{region 'Documentation'}
(*!
<summary>Number of occupied entries.</summary>
*)
{endregion}
{attribute 'monitoring' := 'call'}
PROPERTY PUBLIC ChildCount : UINT //! Number of occupied entries.
GET
ChildCount := FCount;
END_GET
END_PROPERTY

{region 'Documentation'}
(*!
<summary>Records the original array index and returns only registered entries; never invokes a child.</summary>
*)
{endregion}
METHOD PUBLIC GetChild : I_Orchestratable //! Copied child interface at the original occupied index; zero and a latched InvalidAccess for an invalid index.
VAR_INPUT
    Index : DINT; //! Original array index to record and resolve within the occupied prefix.
END_VAR
VAR
    Position : LINT;
END_VAR
GetChild := 0;
IF FReadCount < ReadCapacity THEN
    FReadCount := FReadCount + 1;
    FReadIndices[FReadCount] := Index;
ELSE
    FTraceOverflow := TRUE;
END_IF;

Position := DINT_TO_LINT(Index) - DINT_TO_LINT(FLowerBound) + 1;
IF (Position < 1) OR (Position > UINT_TO_LINT(FCount)) THEN
    FInvalidAccess := TRUE;
    RETURN;
END_IF;
GetChild := FChildren[LINT_TO_UINT(Position)];
END_METHOD

{region 'Documentation'}
(*!
<summary>Copies the fixed registered prefix and clears access evidence without retaining addresses.</summary>
*)
{endregion}
METHOD PUBLIC Initialize : BOOL //! TRUE after copying a valid nonzero occupied prefix; FALSE leaves ChildCount zero.
VAR_INPUT
    Count : UINT; //! Occupied prefix length in 1..ChildCapacity; it must fit the supplied array.
END_VAR
VAR_IN_OUT
    Children : ARRAY[*] OF I_Orchestratable; //! Borrowed array whose occupied interface prefix is copied; keep the referenced children alive.
END_VAR
VAR
    Position : UINT;
    ArrayIndex : DINT;
END_VAR
Initialize := FALSE;
FCount := 0;
FLowerBound := LOWER_BOUND(Children, 1);
FUpperBound := UPPER_BOUND(Children, 1);
FReadCount := 0;
FInvalidAccess := FALSE;
FTraceOverflow := FALSE;
FOR Position := 1 TO ChildCapacity DO
    FChildren[Position] := 0;
END_FOR;
FOR Position := 1 TO ReadCapacity DO
    FReadIndices[Position] := 0;
END_FOR;
IF (Count = 0) OR (Count > ChildCapacity)
    OR (DINT_TO_LINT(FLowerBound) + UINT_TO_LINT(Count) - 1 > DINT_TO_LINT(FUpperBound)) THEN
    RETURN;
END_IF;

FOR Position := 1 TO Count DO
    ArrayIndex := FLowerBound + UINT_TO_DINT(Position) - 1;
    IF Children[ArrayIndex] = 0 THEN
        RETURN;
    END_IF;
    FChildren[Position] := Children[ArrayIndex];
END_FOR;
FCount := Count;
Initialize := TRUE;
END_METHOD

{region 'Documentation'}
(*!
<summary>Latched access outside the registered range.</summary>
*)
{endregion}
{attribute 'monitoring' := 'call'}
PROPERTY PUBLIC InvalidAccess : BOOL //! Latched access outside the registered range.
GET
InvalidAccess := FInvalidAccess;
END_GET
END_PROPERTY

{region 'Documentation'}
(*!
<summary>Number of retained index-access observations.</summary>
*)
{endregion}
{attribute 'monitoring' := 'call'}
PROPERTY PUBLIC ReadCount : UINT //! Number of retained index-access observations.
GET
ReadCount := FReadCount;
END_GET
END_PROPERTY

{region 'Documentation'}
(*!
<summary>Whether the bounded index trace was exhausted.</summary>
*)
{endregion}
{attribute 'monitoring' := 'call'}
PROPERTY PUBLIC TraceOverflow : BOOL //! Whether the bounded index trace was exhausted.
GET
TraceOverflow := FTraceOverflow;
END_GET
END_PROPERTY

END_FUNCTION_BLOCK

// ---- SelfTests/Helper/Orchestration/OrchestrationChildDouble.TcPOU
{region 'Documentation'}
(*!
<summary>Controllable I_Orchestratable boundary for isolated scheduler tests.</summary>
<description>

Stimulus versus commands

The scenario supplies the next ObservationInput at the child FB call after the helper.
Request methods only record invocations; they do not select states or run a copied lifecycle.
This permits independent, explicitly authored normal and exceptional responses.
BeginCycle clears call counters before the helper without changing the prior observation.

Reservation boundary

BeginCycle supplies this cycle's reservation responses, defaulting to Accepted.
Only Accepted sets one local marker; waiting and failure leave it unchanged.
No global publisher or reservation is changed.
The tests verify orchestration call order, not the real owner's budget calculation.
</description>
*)
{endregion}
FUNCTION_BLOCK OrchestrationChildDouble IMPLEMENTS I_Orchestratable
VAR_INPUT
    ObservationInput : ST_OrchestrationObservation; //! Scripted view accepted only when this concrete child body is called.
END_VAR
VAR
    FName : STRING(GVL_Constants.NameLength);
    FExecutionSlot : UINT;
    FInitialized : BOOL;
    FObservation : ST_OrchestrationObservation;
    FCalls : ST_OrchestrationCalls;
    FReservedEntryCount : UINT;
    FExecutionReservationResult : E_EventReservationResult := E_EventReservationResult.Accepted;
    FResetReservationResult : E_EventReservationResult := E_EventReservationResult.Accepted;
END_VAR
VAR CONSTANT
    ReservationMarker : UINT := 1;
END_VAR

FCalls.BodyCount := FCalls.BodyCount + 1;
FObservation := ObservationInput;

{region 'Documentation'}
(*!
<summary>Clears call evidence and supplies reservation responses; retains the prior child view and marker.</summary>
*)
{endregion}
METHOD PUBLIC BeginCycle
VAR_INPUT
    ExecutionReservationResult : E_EventReservationResult := E_EventReservationResult.Accepted; //! Execution admission response for this cycle; Accepted sets the local marker.
    ResetReservationResult : E_EventReservationResult := E_EventReservationResult.Accepted; //! Reset admission response for this cycle; Accepted sets the local marker.
END_VAR
VAR
    EmptyCalls : ST_OrchestrationCalls;
END_VAR
FCalls := EmptyCalls;
FExecutionReservationResult := ExecutionReservationResult;
FResetReservationResult := ResetReservationResult;
END_METHOD

{region 'Documentation'}
(*!
<summary>Interface-call evidence for the current fixture cycle.</summary>
*)
{endregion}
{attribute 'monitoring' := 'variable'}
PROPERTY PUBLIC Calls : ST_OrchestrationCalls //! Interface-call evidence for the current fixture cycle.
GET
Calls := FCalls;
END_GET
END_PROPERTY

{region 'Documentation'}
(*!
<summary>Registration slot retained independently of cyclic observations.</summary>
*)
{endregion}
{attribute 'monitoring' := 'call'}
PROPERTY PUBLIC ExecutionSlot : UINT //! Registration slot retained independently of cyclic observations.
GET
ExecutionSlot := FExecutionSlot;
END_GET
SET
FExecutionSlot := ExecutionSlot;
END_SET
END_PROPERTY

{region 'Documentation'}
(*!
<summary>Releases only the local marker and records the released amount; repeated calls are idempotent.</summary>
*)
{endregion}
METHOD PUBLIC FreeReservedEvents : BOOL //! Always TRUE after clearing the local marker; the call and released amount remain recorded.
FCalls.FreeCount := FCalls.FreeCount + 1;
FCalls.ReleasedEntryCount := FCalls.ReleasedEntryCount + FReservedEntryCount;
FReservedEntryCount := 0;
FreeReservedEvents := TRUE;
END_METHOD

{region 'Documentation'}
(*!
<summary>Scripted child failure classification.</summary>
*)
{endregion}
{attribute 'monitoring' := 'call'}
PROPERTY PUBLIC HasError : BOOL //! Scripted child failure classification.
GET
HasError := FObservation.Result = E_Result.Error;
END_GET
END_PROPERTY

{region 'Documentation'}
(*!
<summary>Resets the local interface double; it has no timers, publisher or production lifecycle.</summary>
*)
{endregion}
METHOD PUBLIC Initialize
VAR_INPUT
    Name : STRING(GVL_Constants.NameLength); //! Diagnostic child name retained by the fixture.
    Slot : UINT; //! Registered execution slot retained independently of scripted observations.
END_VAR
VAR
    EmptyCalls : ST_OrchestrationCalls;
    InitialView : ST_OrchestrationObservation;
END_VAR
FName := Name;
FExecutionSlot := Slot;
FObservation := InitialView;
FCalls := EmptyCalls;
FReservedEntryCount := 0;
FExecutionReservationResult := E_EventReservationResult.Accepted;
FResetReservationResult := E_EventReservationResult.Accepted;
FInitialized := TRUE;
END_METHOD

{region 'Documentation'}
(*!
<summary>Scripted terminal completion signal.</summary>
*)
{endregion}
{attribute 'monitoring' := 'call'}
PROPERTY PUBLIC IsComplete : BOOL //! Scripted terminal completion signal.
GET
IsComplete := FObservation.Complete;
END_GET
END_PROPERTY

{region 'Documentation'}
(*!
<summary>Whether the double has been explicitly configured.</summary>
*)
{endregion}
{attribute 'monitoring' := 'call'}
PROPERTY PUBLIC IsInitialized : BOOL //! Whether the double has been explicitly configured.
GET
IsInitialized := FInitialized;
END_GET
END_PROPERTY

{region 'Documentation'}
(*!
<summary>Scripted readiness, independent of helper requests.</summary>
*)
{endregion}
{attribute 'monitoring' := 'call'}
PROPERTY PUBLIC IsReady : BOOL //! Scripted readiness, independent of helper requests.
GET
IsReady := FObservation.Ready;
END_GET
END_PROPERTY

{region 'Documentation'}
(*!
<summary>Diagnostic child identity.</summary>
*)
{endregion}
{attribute 'monitoring' := 'variable'}
PROPERTY PUBLIC Name : STRING(GVL_Constants.NameLength) //! Diagnostic child identity.
GET
Name := FName;
END_GET
END_PROPERTY

{region 'Documentation'}
(*!
<summary>Current scripted snapshot; requests cannot change it.</summary>
*)
{endregion}
{attribute 'monitoring' := 'variable'}
PROPERTY PUBLIC Observation : ST_OrchestrationObservation //! Current scripted snapshot; requests cannot change it.
GET
Observation := FObservation;
END_GET
END_PROPERTY

{region 'Documentation'}
(*!
<summary>Records the Abort request without changing the scripted state.</summary>
*)
{endregion}
METHOD PUBLIC RequestAbort
FCalls.AbortCount := FCalls.AbortCount + 1;
END_METHOD

{region 'Documentation'}
(*!
<summary>Records the Reset request without changing the scripted state.</summary>
*)
{endregion}
METHOD PUBLIC RequestReset
FCalls.ResetCount := FCalls.ResetCount + 1;

FCalls.ResetWithoutReservation := FCalls.ResetWithoutReservation OR (FReservedEntryCount = 0);
END_METHOD

{region 'Documentation'}
(*!
<summary>Records the Start request without changing the scripted state.</summary>
*)
{endregion}
METHOD PUBLIC RequestStart
FCalls.StartCount := FCalls.StartCount + 1;
FCalls.StartWithoutReservation := FCalls.StartWithoutReservation OR (FReservedEntryCount = 0);
END_METHOD

{region 'Documentation'}
(*!
<summary>Local admission marker, not a global Event Buffer contribution.</summary>
*)
{endregion}
{attribute 'monitoring' := 'call'}
PROPERTY PUBLIC ReservedEntryCount : UINT //! Local admission marker, not a global Event Buffer contribution.
GET
ReservedEntryCount := FReservedEntryCount;
END_GET
END_PROPERTY

{region 'Documentation'}
(*!
<summary>Returns the scripted execution admission response; only Accepted sets the local marker.</summary>
*)
{endregion}
METHOD PUBLIC ReserveExecutionEvents : E_EventReservationResult //! Scripted execution admission response; only Accepted installs the local marker.
FCalls.ExecutionReservationCount := FCalls.ExecutionReservationCount + 1;
IF FExecutionReservationResult = E_EventReservationResult.Accepted THEN
    FReservedEntryCount := ReservationMarker;
END_IF;
ReserveExecutionEvents := FExecutionReservationResult;
END_METHOD

{region 'Documentation'}
(*!
<summary>Returns the scripted reset admission response; only Accepted sets the local marker.</summary>
*)
{endregion}
METHOD PUBLIC ReserveResetEvents : E_EventReservationResult //! Scripted Reset admission response; only Accepted installs the local marker.
FCalls.ResetReservationCount := FCalls.ResetReservationCount + 1;
IF FResetReservationResult = E_EventReservationResult.Accepted THEN
    FReservedEntryCount := ReservationMarker;
END_IF;
ReserveResetEvents := FResetReservationResult;
END_METHOD

{region 'Documentation'}
(*!
<summary>Scripted child result.</summary>
*)
{endregion}
{attribute 'monitoring' := 'call'}
PROPERTY PUBLIC Result : E_Result //! Scripted child result.
GET
Result := FObservation.Result;
END_GET
END_PROPERTY

{region 'Documentation'}
(*!
<summary>View applied on the most recent child call.</summary>
*)
{endregion}
{attribute 'monitoring' := 'call'}
PROPERTY PUBLIC State : E_State //! View applied on the most recent child call.
GET
State := FObservation.State;
END_GET
END_PROPERTY

END_FUNCTION_BLOCK

// ---- SelfTests/TestCases/TestSuite_Orchestrator/Test_OrchestratorNegativeBounds.TcPOU
{region 'Documentation'}
(*!
<summary>Checks the same execution trace with actual indices -3 through -1.</summary>
*)
{endregion}
FUNCTION_BLOCK Test_OrchestratorNegativeBounds EXTENDS OrchestrationTestBase

SUPER^();

{region 'Documentation'}
(*!
<summary>Defines this scenario independently of the subject's internal fields.</summary>
*)
{endregion}
METHOD PROTECTED ConfigureScenario
FArrayLayout := E_OrchestrationArrayLayout.Negative;
FChildCount := 3;
ConfigureStandardSequence();
END_METHOD

END_FUNCTION_BLOCK

// ---- SelfTests/TestCases/TestSuite_Orchestrator/Test_OrchestratorUnusedCapacity.TcPOU
{region 'Documentation'}
(*!
<summary>Checks that unused array capacity at indices 4 through 6 is never processed.</summary>
*)
{endregion}
FUNCTION_BLOCK Test_OrchestratorUnusedCapacity EXTENDS OrchestrationTestBase

SUPER^();

{region 'Documentation'}
(*!
<summary>Defines this scenario independently of the subject's internal fields.</summary>
*)
{endregion}
METHOD PROTECTED ConfigureScenario
FArrayLayout := E_OrchestrationArrayLayout.SpareCapacity;
FChildCount := 3;
ConfigureStandardSequence();
END_METHOD

END_FUNCTION_BLOCK

// ---- SelfTests/TestCases/TestSuite_Orchestrator/Test_OrchestratorSingleChild.TcPOU
{region 'Documentation'}
(*!
<summary>Checks a single registered child without a successor or unused-capacity access.</summary>
*)
{endregion}
FUNCTION_BLOCK Test_OrchestratorSingleChild EXTENDS OrchestrationTestBase

SUPER^();

{region 'Documentation'}
(*!
<summary>Defines this scenario independently of the subject's internal fields.</summary>
*)
{endregion}
METHOD PROTECTED ConfigureScenario
FArrayLayout := E_OrchestrationArrayLayout.Ordinary;
FChildCount := 1;
FStepCount := 4;

{region "Cycle 01 - Idle readiness"}
FSteps[1].Task := E_OrchestratorTask.Idle;
FSteps[1].ExpectedReady := TRUE;
{endregion}

{region "Cycle 02 - Start child 1"}
FSteps[2].Children[1].State := E_State.Completed;
FSteps[2].Children[1].Ready := FALSE;
FSteps[2].Children[1].Complete := TRUE;
FSteps[2].Children[1].Result := E_Result.Passed;
FSteps[2].ExpectedStartChild := 1;
FSteps[2].ExpectedSlot := 1;
FSteps[2].ExpectedReservations[1] := 1;
{endregion}

{region "Cycle 03 - Completed observation"}
FSteps[3].Children[1].State := E_State.Completed;
FSteps[3].Children[1].Ready := FALSE;
FSteps[3].Children[1].Complete := TRUE;
FSteps[3].Children[1].Result := E_Result.Passed;
FSteps[3].ExpectedReleasedEntries[1] := 1;
FSteps[3].ExpectedFinished := TRUE;
{endregion}

{region "Cycle 04 - Completed observation"}
FSteps[4].Children[1].State := E_State.Completed;
FSteps[4].Children[1].Ready := FALSE;
FSteps[4].Children[1].Complete := TRUE;
FSteps[4].Children[1].Result := E_Result.Passed;
FSteps[4].ExpectedFinished := TRUE;
{endregion}
END_METHOD

END_FUNCTION_BLOCK

// ---- SelfTests/TestCases/TestSuite_Orchestrator/Test_OrchestratorIdleReadiness.TcPOU
{region 'Documentation'}
(*!
<summary>Checks that readiness follows prior child observations and recovers without dispatch or diagnostics.</summary>
*)
{endregion}
FUNCTION_BLOCK Test_OrchestratorIdleReadiness EXTENDS OrchestrationTestBase

SUPER^();

{region 'Documentation'}
(*!
<summary>Defines independent stimuli and expected requests, reservations, task status and diagnostic counts.</summary>
*)
{endregion}
METHOD PROTECTED ConfigureScenario
FStepCount := 4;

{region "01 - Make the second child not ready after helper observation"}
FSteps[1].Task := E_OrchestratorTask.Idle;
FSteps[1].Children[2].Ready := FALSE;
FSteps[1].ExpectedReady := TRUE;
{endregion}

{region "02 - Observe not-ready child without dispatch"}
FSteps[2].Task := E_OrchestratorTask.Idle;
FSteps[2].Children[2].Ready := FALSE;
{endregion}

{region "03 - Restore child readiness after this observation"}
FSteps[3].Task := E_OrchestratorTask.Idle;
{endregion}

{region "04 - Observe restored readiness"}
FSteps[4].Task := E_OrchestratorTask.Idle;
FSteps[4].ExpectedReady := TRUE;
{endregion}
END_METHOD

END_FUNCTION_BLOCK

// ---- SelfTests/TestCases/TestSuite_Orchestrator/Test_OrchestratorMissingStartReaction.TcPOU
{region 'Documentation'}
(*!
<summary>Detects missing Start response on the following call, releases its reservation and prevents retries.</summary>
*)
{endregion}
FUNCTION_BLOCK Test_OrchestratorMissingStartReaction EXTENDS OrchestrationTestBase

SUPER^();

{region 'Documentation'}
(*!
<summary>Defines independent stimuli and expected requests, reservations, task status and diagnostic counts.</summary>
*)
{endregion}
METHOD PROTECTED ConfigureScenario
FStepCount := 12;

{region "01 - Idle readiness before child processing"}
FSteps[1].Task := E_OrchestratorTask.Idle;
FSteps[1].ExpectedReady := TRUE;
{endregion}

{region "02 - Request Start but leave child Idle"}
FSteps[2].ExpectedStartChild := 1;
FSteps[2].ExpectedSlot := 1;
FSteps[2].ExpectedReservations[1] := 1;
{endregion}

{region "03 - Following helper call must reject missing response"}
FSteps[3].ExpectedSlot := 1;
FSteps[3].ExpectedDiagnosticCount := 1;
FSteps[3].ExpectedReleasedEntries[1] := 1;
FSteps[3].ExpectedResult := E_Result.Error;
{endregion}

{region "04 - No retry or duplicate diagnostic"}
FSteps[4].ExpectedSlot := 1;
FSteps[4].ExpectedDiagnosticCount := 1;
FSteps[4].ExpectedResult := E_Result.Error;
{endregion}

{region "05 - Idle preserves the held error"}
FSteps[5].Task := E_OrchestratorTask.Idle;
FSteps[5].ExpectedDiagnosticCount := 1;
FSteps[5].ExpectedResult := E_Result.Error;
{endregion}

{region "06 - Execution cannot bypass held error"}
FSteps[6].ExpectedDiagnosticCount := 1;
FSteps[6].ExpectedResult := E_Result.Error;
{endregion}

{region "07 - New Reset clears helper error without clearing captured evidence"}
FSteps[7].Task := E_OrchestratorTask.Reset;
FSteps[7].ExpectedDiagnosticCount := 1;
{endregion}

{region "08 - All already-ready children count as reset-complete"}
FSteps[8].Task := E_OrchestratorTask.Reset;
FSteps[8].ExpectedDiagnosticCount := 1;
FSteps[8].ExpectedResetFinished := TRUE;
{endregion}

{region "09 - Owner returns to ready Idle"}
FSteps[9].Task := E_OrchestratorTask.Idle;
FSteps[9].ExpectedDiagnosticCount := 1;
FSteps[9].ExpectedReady := TRUE;
{endregion}

{region "10 - Start is admitted again only after Reset"}
FSteps[10].Children[1].State := E_State.Completed;
FSteps[10].Children[1].Result := E_Result.Passed;
FSteps[10].Children[1].Ready := FALSE;
FSteps[10].Children[1].Complete := TRUE;
FSteps[10].ExpectedStartChild := 1;
FSteps[10].ExpectedSlot := 1;
FSteps[10].ExpectedDiagnosticCount := 1;
FSteps[10].ExpectedReservations[1] := 1;
{endregion}

{region "11 - Successful start response does not create another diagnostic"}
FSteps[11].Children[1].State := E_State.Completed;
FSteps[11].Children[1].Result := E_Result.Passed;
FSteps[11].Children[1].Ready := FALSE;
FSteps[11].Children[1].Complete := TRUE;
FSteps[11].ExpectedSlot := 2;
FSteps[11].ExpectedDiagnosticCount := 1;
FSteps[11].ExpectedReleasedEntries[1] := 1;
{endregion}

{region "12 - Owner stops the local scenario without starting later children"}
FSteps[12].Task := E_OrchestratorTask.Idle;
FSteps[12].Children[1].State := E_State.Completed;
FSteps[12].Children[1].Result := E_Result.Passed;
FSteps[12].Children[1].Ready := FALSE;
FSteps[12].Children[1].Complete := TRUE;
FSteps[12].ExpectedDiagnosticCount := 1;
{endregion}
END_METHOD

END_FUNCTION_BLOCK

// ---- SelfTests/TestCases/TestSuite_Orchestrator/Test_OrchestratorChildError.TcPOU
{region 'Documentation'}
(*!
<summary>Holds a child Error, prevents subsequent Starts and releases only after terminal observation.</summary>
*)
{endregion}
FUNCTION_BLOCK Test_OrchestratorChildError EXTENDS OrchestrationTestBase

SUPER^();

{region 'Documentation'}
(*!
<summary>Defines independent stimuli and expected requests, reservations, task status and diagnostic counts.</summary>
*)
{endregion}
METHOD PROTECTED ConfigureScenario
FStepCount := 8;

{region "01 - Idle readiness before child processing"}
FSteps[1].Task := E_OrchestratorTask.Idle;
FSteps[1].ExpectedReady := TRUE;
{endregion}

{region "02 - Start first child"}
FSteps[2].Children[1].State := E_State.Running;
FSteps[2].Children[1].Ready := FALSE;
FSteps[2].ExpectedStartChild := 1;
FSteps[2].ExpectedSlot := 1;
FSteps[2].ExpectedReservations[1] := 1;
{endregion}

{region "03 - Child reports Error after helper call"}
FSteps[3].Children[1].State := E_State.Running;
FSteps[3].Children[1].Result := E_Result.Error;
FSteps[3].Children[1].Ready := FALSE;
FSteps[3].ExpectedSlot := 1;
FSteps[3].ExpectedReservations[1] := 1;
{endregion}

{region "04 - Observe Error and retain active reservation"}
FSteps[4].Children[1].State := E_State.Running;
FSteps[4].Children[1].Result := E_Result.Error;
FSteps[4].Children[1].Ready := FALSE;
FSteps[4].ExpectedSlot := 1;
FSteps[4].ExpectedDiagnosticCount := 1;
FSteps[4].ExpectedReservations[1] := 1;
FSteps[4].ExpectedResult := E_Result.Error;
{endregion}

{region "05 - Failing child reaches terminal state"}
FSteps[5].Children[1].State := E_State.Completed;
FSteps[5].Children[1].Result := E_Result.Error;
FSteps[5].Children[1].Ready := FALSE;
FSteps[5].Children[1].Complete := TRUE;
FSteps[5].ExpectedSlot := 1;
FSteps[5].ExpectedDiagnosticCount := 1;
FSteps[5].ExpectedReservations[1] := 1;
FSteps[5].ExpectedResult := E_Result.Error;
{endregion}

{region "06 - Release terminal reservation without advancing execution"}
FSteps[6].Children[1].State := E_State.Completed;
FSteps[6].Children[1].Result := E_Result.Error;
FSteps[6].Children[1].Ready := FALSE;
FSteps[6].Children[1].Complete := TRUE;
FSteps[6].ExpectedSlot := 1;
FSteps[6].ExpectedDiagnosticCount := 1;
FSteps[6].ExpectedReleasedEntries[1] := 1;
FSteps[6].ExpectedResult := E_Result.Error;
{endregion}

{region "07 - Idle must not clear Error"}
FSteps[7].Task := E_OrchestratorTask.Idle;
FSteps[7].Children[1].State := E_State.Completed;
FSteps[7].Children[1].Result := E_Result.Error;
FSteps[7].Children[1].Ready := FALSE;
FSteps[7].Children[1].Complete := TRUE;
FSteps[7].ExpectedDiagnosticCount := 1;
FSteps[7].ExpectedResult := E_Result.Error;
{endregion}

{region "08 - Repeated Idle remains quiet"}
FSteps[8].Task := E_OrchestratorTask.Idle;
FSteps[8].Children[1].State := E_State.Completed;
FSteps[8].Children[1].Result := E_Result.Error;
FSteps[8].Children[1].Ready := FALSE;
FSteps[8].Children[1].Complete := TRUE;
FSteps[8].ExpectedDiagnosticCount := 1;
FSteps[8].ExpectedResult := E_Result.Error;
{endregion}
END_METHOD

END_FUNCTION_BLOCK

// ---- SelfTests/TestCases/TestSuite_Orchestrator/Test_OrchestratorUnexpectedAbort.TcPOU
{region 'Documentation'}
(*!
<summary>Treats a subordinate Abort during execution as a helper Error rather than normal completion.</summary>
*)
{endregion}
FUNCTION_BLOCK Test_OrchestratorUnexpectedAbort EXTENDS OrchestrationTestBase

SUPER^();

{region 'Documentation'}
(*!
<summary>Defines independent stimuli and expected requests, reservations, task status and diagnostic counts.</summary>
*)
{endregion}
METHOD PROTECTED ConfigureScenario
FStepCount := 6;

{region "01 - Idle readiness before child processing"}
FSteps[1].Task := E_OrchestratorTask.Idle;
FSteps[1].ExpectedReady := TRUE;
{endregion}

{region "02 - Start first child"}
FSteps[2].Children[1].State := E_State.Running;
FSteps[2].Children[1].Ready := FALSE;
FSteps[2].ExpectedStartChild := 1;
FSteps[2].ExpectedSlot := 1;
FSteps[2].ExpectedReservations[1] := 1;
{endregion}

{region "03 - Child reports unexpected Abort"}
FSteps[3].Children[1].State := E_State.Running;
FSteps[3].Children[1].Result := E_Result.Abort;
FSteps[3].Children[1].Ready := FALSE;
FSteps[3].ExpectedSlot := 1;
FSteps[3].ExpectedReservations[1] := 1;
{endregion}

{region "04 - Observe unexpected Abort while child finishes"}
FSteps[4].Children[1].State := E_State.Completed;
FSteps[4].Children[1].Result := E_Result.Abort;
FSteps[4].Children[1].Ready := FALSE;
FSteps[4].Children[1].Complete := TRUE;
FSteps[4].ExpectedSlot := 1;
FSteps[4].ExpectedDiagnosticCount := 1;
FSteps[4].ExpectedReservations[1] := 1;
FSteps[4].ExpectedResult := E_Result.Error;
{endregion}

{region "05 - Release without starting the successor"}
FSteps[5].Children[1].State := E_State.Completed;
FSteps[5].Children[1].Result := E_Result.Abort;
FSteps[5].Children[1].Ready := FALSE;
FSteps[5].Children[1].Complete := TRUE;
FSteps[5].ExpectedSlot := 1;
FSteps[5].ExpectedDiagnosticCount := 1;
FSteps[5].ExpectedReleasedEntries[1] := 1;
FSteps[5].ExpectedResult := E_Result.Error;
{endregion}

{region "06 - Held Error prevents a later Start"}
FSteps[6].Children[1].State := E_State.Completed;
FSteps[6].Children[1].Result := E_Result.Abort;
FSteps[6].Children[1].Ready := FALSE;
FSteps[6].Children[1].Complete := TRUE;
FSteps[6].ExpectedSlot := 1;
FSteps[6].ExpectedDiagnosticCount := 1;
FSteps[6].ExpectedResult := E_Result.Error;
{endregion}
END_METHOD

END_FUNCTION_BLOCK

// ---- SelfTests/TestCases/TestSuite_Orchestrator/Test_OrchestratorAbortInterruption.TcPOU
{region 'Documentation'}
(*!
<summary>Changes the owner task to Abort, requests only the active child and observes terminal cleanup.</summary>
*)
{endregion}
FUNCTION_BLOCK Test_OrchestratorAbortInterruption EXTENDS OrchestrationTestBase

SUPER^();

{region 'Documentation'}
(*!
<summary>Defines independent stimuli and expected requests, reservations, task status and diagnostic counts.</summary>
*)
{endregion}
METHOD PROTECTED ConfigureScenario
FStepCount := 8;

{region "01 - Idle readiness before child processing"}
FSteps[1].Task := E_OrchestratorTask.Idle;
FSteps[1].ExpectedReady := TRUE;
{endregion}

{region "02 - Start first child"}
FSteps[2].Children[1].State := E_State.Running;
FSteps[2].Children[1].Ready := FALSE;
FSteps[2].ExpectedStartChild := 1;
FSteps[2].ExpectedSlot := 1;
FSteps[2].ExpectedReservations[1] := 1;
{endregion}

{region "03 - Abort replaces Execution in the same helper call"}
FSteps[3].Task := E_OrchestratorTask.Abort;
FSteps[3].Children[1].State := E_State.Aborting;
FSteps[3].Children[1].Result := E_Result.Abort;
FSteps[3].Children[1].Ready := FALSE;
FSteps[3].ExpectedReservations[1] := 1;
FSteps[3].ExpectedAbortRequests[1] := 1;
{endregion}

{region "04 - Already-aborting child receives no duplicate request"}
FSteps[4].Task := E_OrchestratorTask.Abort;
FSteps[4].Children[1].State := E_State.Aborting;
FSteps[4].Children[1].Result := E_Result.Abort;
FSteps[4].Children[1].Ready := FALSE;
FSteps[4].ExpectedReservations[1] := 1;
{endregion}

{region "05 - Child reaches Completed with Abort"}
FSteps[5].Task := E_OrchestratorTask.Abort;
FSteps[5].Children[1].State := E_State.Completed;
FSteps[5].Children[1].Result := E_Result.Abort;
FSteps[5].Children[1].Ready := FALSE;
FSteps[5].Children[1].Complete := TRUE;
FSteps[5].ExpectedReservations[1] := 1;
{endregion}

{region "06 - Observe Abort completion and release"}
FSteps[6].Task := E_OrchestratorTask.Abort;
FSteps[6].Children[1].State := E_State.Completed;
FSteps[6].Children[1].Result := E_Result.Abort;
FSteps[6].Children[1].Ready := FALSE;
FSteps[6].Children[1].Complete := TRUE;
FSteps[6].ExpectedReleasedEntries[1] := 1;
FSteps[6].ExpectedAbortFinished := TRUE;
{endregion}

{region "07 - Completion does not select Idle autonomously"}
FSteps[7].Task := E_OrchestratorTask.Abort;
FSteps[7].Children[1].State := E_State.Completed;
FSteps[7].Children[1].Result := E_Result.Abort;
FSteps[7].Children[1].Ready := FALSE;
FSteps[7].Children[1].Complete := TRUE;
FSteps[7].ExpectedAbortFinished := TRUE;
{endregion}

{region "08 - Owner explicitly selects Idle"}
FSteps[8].Task := E_OrchestratorTask.Idle;
FSteps[8].Children[1].State := E_State.Completed;
FSteps[8].Children[1].Result := E_Result.Abort;
FSteps[8].Children[1].Ready := FALSE;
FSteps[8].Children[1].Complete := TRUE;
{endregion}
END_METHOD

END_FUNCTION_BLOCK

// ---- SelfTests/TestCases/TestSuite_Orchestrator/Test_OrchestratorIdleInterruption.TcPOU
{region 'Documentation'}
(*!
<summary>Idle stops new dispatch without forcing child Abort or releasing an unfinished reservation.</summary>
*)
{endregion}
FUNCTION_BLOCK Test_OrchestratorIdleInterruption EXTENDS OrchestrationTestBase

SUPER^();

{region 'Documentation'}
(*!
<summary>Defines independent stimuli and expected requests, reservations, task status and diagnostic counts.</summary>
*)
{endregion}
METHOD PROTECTED ConfigureScenario
FStepCount := 6;

{region "01 - Idle readiness before child processing"}
FSteps[1].Task := E_OrchestratorTask.Idle;
FSteps[1].ExpectedReady := TRUE;
{endregion}

{region "02 - Start first child"}
FSteps[2].Children[1].State := E_State.Running;
FSteps[2].Children[1].Ready := FALSE;
FSteps[2].ExpectedStartChild := 1;
FSteps[2].ExpectedSlot := 1;
FSteps[2].ExpectedReservations[1] := 1;
{endregion}

{region "03 - Idle leaves running child and reservation intact"}
FSteps[3].Task := E_OrchestratorTask.Idle;
FSteps[3].Children[1].State := E_State.Running;
FSteps[3].Children[1].Ready := FALSE;
FSteps[3].ExpectedReservations[1] := 1;
{endregion}

{region "04 - Child finishes while owner remains Idle"}
FSteps[4].Task := E_OrchestratorTask.Idle;
FSteps[4].Children[1].State := E_State.Completed;
FSteps[4].Children[1].Result := E_Result.Passed;
FSteps[4].Children[1].Ready := FALSE;
FSteps[4].Children[1].Complete := TRUE;
FSteps[4].ExpectedReservations[1] := 1;
{endregion}

{region "05 - Idle releases the finished child only"}
FSteps[5].Task := E_OrchestratorTask.Idle;
FSteps[5].Children[1].State := E_State.Completed;
FSteps[5].Children[1].Result := E_Result.Passed;
FSteps[5].Children[1].Ready := FALSE;
FSteps[5].Children[1].Complete := TRUE;
FSteps[5].ExpectedReleasedEntries[1] := 1;
{endregion}

{region "06 - Idle does not start the next child"}
FSteps[6].Task := E_OrchestratorTask.Idle;
FSteps[6].Children[1].State := E_State.Completed;
FSteps[6].Children[1].Result := E_Result.Passed;
FSteps[6].Children[1].Ready := FALSE;
FSteps[6].Children[1].Complete := TRUE;
{endregion}
END_METHOD

END_FUNCTION_BLOCK

// ---- SelfTests/TestCases/TestSuite_Orchestrator/Test_OrchestratorResetInterruption.TcPOU
{region 'Documentation'}
(*!
<summary>Reset replaces Execution and may dispatch subsequent child resets before prior reset completion.</summary>
*)
{endregion}
FUNCTION_BLOCK Test_OrchestratorResetInterruption EXTENDS OrchestrationTestBase

SUPER^();

{region 'Documentation'}
(*!
<summary>Defines independent stimuli and expected requests, reservations, task status and diagnostic counts.</summary>
*)
{endregion}
METHOD PROTECTED ConfigureScenario
FStepCount := 10;

{region "01 - Idle readiness before child processing"}
FSteps[1].Task := E_OrchestratorTask.Idle;
FSteps[1].ExpectedReady := TRUE;
{endregion}

{region "02 - Execution begins; other resources become not ready"}
FSteps[2].Children[1].State := E_State.Running;
FSteps[2].Children[1].Ready := FALSE;
FSteps[2].Children[2].Ready := FALSE;
FSteps[2].Children[3].Ready := FALSE;
FSteps[2].ExpectedStartChild := 1;
FSteps[2].ExpectedSlot := 1;
FSteps[2].ExpectedReservations[1] := 1;
{endregion}

{region "03 - Reset first child in the task-entry call"}
FSteps[3].Task := E_OrchestratorTask.Reset;
FSteps[3].Children[1].State := E_State.Reset;
FSteps[3].Children[1].Ready := FALSE;
FSteps[3].Children[2].Ready := FALSE;
FSteps[3].Children[3].Ready := FALSE;
FSteps[3].ExpectedResetChild := 1;
FSteps[3].ExpectedReservations[1] := 1;
{endregion}

{region "04 - Dispatch second Reset while first is still active"}
FSteps[4].Task := E_OrchestratorTask.Reset;
FSteps[4].Children[1].State := E_State.Reset;
FSteps[4].Children[1].Ready := FALSE;
FSteps[4].Children[2].State := E_State.Reset;
FSteps[4].Children[2].Ready := FALSE;
FSteps[4].Children[3].Ready := FALSE;
FSteps[4].ExpectedResetChild := 2;
FSteps[4].ExpectedReservations[1] := 1;
FSteps[4].ExpectedReservations[2] := 1;
{endregion}

{region "05 - Dispatch third Reset; first finishes afterwards"}
FSteps[5].Task := E_OrchestratorTask.Reset;
FSteps[5].Children[2].State := E_State.Reset;
FSteps[5].Children[2].Ready := FALSE;
FSteps[5].Children[3].State := E_State.Reset;
FSteps[5].Children[3].Ready := FALSE;
FSteps[5].ExpectedResetChild := 3;
FSteps[5].ExpectedReservations[1] := 1;
FSteps[5].ExpectedReservations[2] := 1;
FSteps[5].ExpectedReservations[3] := 1;
{endregion}

{region "06 - Release first; second finishes afterwards"}
FSteps[6].Task := E_OrchestratorTask.Reset;
FSteps[6].Children[3].State := E_State.Reset;
FSteps[6].Children[3].Ready := FALSE;
FSteps[6].ExpectedReservations[2] := 1;
FSteps[6].ExpectedReservations[3] := 1;
FSteps[6].ExpectedReleasedEntries[1] := 1;
{endregion}

{region "07 - Release second; third finishes afterwards"}
FSteps[7].Task := E_OrchestratorTask.Reset;
FSteps[7].ExpectedReservations[3] := 1;
FSteps[7].ExpectedReleasedEntries[2] := 1;
{endregion}

{region "08 - All reset observations are ready and reconciled"}
FSteps[8].Task := E_OrchestratorTask.Reset;
FSteps[8].ExpectedReleasedEntries[3] := 1;
FSteps[8].ExpectedResetFinished := TRUE;
{endregion}

{region "09 - Repeated Reset task does not restart dispatch"}
FSteps[9].Task := E_OrchestratorTask.Reset;
FSteps[9].ExpectedResetFinished := TRUE;
{endregion}

{region "10 - Only owner task change makes helper ready"}
FSteps[10].Task := E_OrchestratorTask.Idle;
FSteps[10].ExpectedReady := TRUE;
{endregion}
END_METHOD

END_FUNCTION_BLOCK

// ---- SelfTests/TestCases/TestSuite_Orchestrator/Test_OrchestratorResetContinuesAfterError.TcPOU
{region 'Documentation'}
(*!
<summary>Reset ignores unprocessed stale results, retains processed child errors and still attempts every child.</summary>
*)
{endregion}
FUNCTION_BLOCK Test_OrchestratorResetContinuesAfterError EXTENDS OrchestrationTestBase

SUPER^();

{region 'Documentation'}
(*!
<summary>Defines independent stimuli and expected requests, reservations, task status and diagnostic counts.</summary>
*)
{endregion}
METHOD PROTECTED ConfigureScenario
FStepCount := 8;

{region "01 - Establish previous terminal results through child calls"}
FSteps[1].Task := E_OrchestratorTask.Idle;
FSteps[1].Children[1].State := E_State.Completed;
FSteps[1].Children[1].Result := E_Result.Passed;
FSteps[1].Children[1].Ready := FALSE;
FSteps[1].Children[1].Complete := TRUE;
FSteps[1].Children[2].State := E_State.Completed;
FSteps[1].Children[2].Result := E_Result.Error;
FSteps[1].Children[2].Ready := FALSE;
FSteps[1].Children[2].Complete := TRUE;
FSteps[1].Children[3].State := E_State.Completed;
FSteps[1].Children[3].Result := E_Result.Passed;
FSteps[1].Children[3].Ready := FALSE;
FSteps[1].Children[3].Complete := TRUE;
FSteps[1].ExpectedReady := TRUE;
{endregion}

{region "02 - Reset first; ignore old Error in not-yet-reset second child"}
FSteps[2].Task := E_OrchestratorTask.Reset;
FSteps[2].Children[1].State := E_State.Completed;
FSteps[2].Children[1].Result := E_Result.Error;
FSteps[2].Children[1].Ready := FALSE;
FSteps[2].Children[1].Complete := TRUE;
FSteps[2].Children[2].State := E_State.Completed;
FSteps[2].Children[2].Result := E_Result.Error;
FSteps[2].Children[2].Ready := FALSE;
FSteps[2].Children[2].Complete := TRUE;
FSteps[2].Children[3].State := E_State.Completed;
FSteps[2].Children[3].Result := E_Result.Passed;
FSteps[2].Children[3].Ready := FALSE;
FSteps[2].Children[3].Complete := TRUE;
FSteps[2].ExpectedResetChild := 1;
FSteps[2].ExpectedReservations[1] := 1;
{endregion}

{region "03 - First Reset failed; still dispatch second"}
FSteps[3].Task := E_OrchestratorTask.Reset;
FSteps[3].Children[1].State := E_State.Completed;
FSteps[3].Children[1].Result := E_Result.Error;
FSteps[3].Children[1].Ready := FALSE;
FSteps[3].Children[1].Complete := TRUE;
FSteps[3].Children[2].State := E_State.Reset;
FSteps[3].Children[2].Ready := FALSE;
FSteps[3].Children[3].State := E_State.Completed;
FSteps[3].Children[3].Result := E_Result.Passed;
FSteps[3].Children[3].Ready := FALSE;
FSteps[3].Children[3].Complete := TRUE;
FSteps[3].ExpectedResetChild := 2;
FSteps[3].ExpectedDiagnosticCount := 1;
FSteps[3].ExpectedReservations[1] := 1;
FSteps[3].ExpectedReservations[2] := 1;
FSteps[3].ExpectedResult := E_Result.Error;
{endregion}

{region "04 - Keep failure while dispatching third"}
FSteps[4].Task := E_OrchestratorTask.Reset;
FSteps[4].Children[1].State := E_State.Completed;
FSteps[4].Children[1].Result := E_Result.Error;
FSteps[4].Children[1].Ready := FALSE;
FSteps[4].Children[1].Complete := TRUE;
FSteps[4].Children[3].State := E_State.Reset;
FSteps[4].Children[3].Ready := FALSE;
FSteps[4].ExpectedResetChild := 3;
FSteps[4].ExpectedDiagnosticCount := 1;
FSteps[4].ExpectedReservations[1] := 1;
FSteps[4].ExpectedReservations[2] := 1;
FSteps[4].ExpectedReservations[3] := 1;
FSteps[4].ExpectedResult := E_Result.Error;
{endregion}

{region "05 - Release successful second Reset"}
FSteps[5].Task := E_OrchestratorTask.Reset;
FSteps[5].Children[1].State := E_State.Completed;
FSteps[5].Children[1].Result := E_Result.Error;
FSteps[5].Children[1].Ready := FALSE;
FSteps[5].Children[1].Complete := TRUE;
FSteps[5].ExpectedDiagnosticCount := 1;
FSteps[5].ExpectedReservations[1] := 1;
FSteps[5].ExpectedReservations[3] := 1;
FSteps[5].ExpectedReleasedEntries[2] := 1;
FSteps[5].ExpectedResult := E_Result.Error;
{endregion}

{region "06 - Failed terminal child counts as finished, not ready"}
FSteps[6].Task := E_OrchestratorTask.Reset;
FSteps[6].Children[1].State := E_State.Completed;
FSteps[6].Children[1].Result := E_Result.Error;
FSteps[6].Children[1].Ready := FALSE;
FSteps[6].Children[1].Complete := TRUE;
FSteps[6].ExpectedDiagnosticCount := 1;
FSteps[6].ExpectedReservations[1] := 1;
FSteps[6].ExpectedReleasedEntries[3] := 1;
FSteps[6].ExpectedResetFinished := TRUE;
FSteps[6].ExpectedResult := E_Result.Error;
{endregion}

{region "07 - Idle reconciles failed terminal child reservation"}
FSteps[7].Task := E_OrchestratorTask.Idle;
FSteps[7].Children[1].State := E_State.Completed;
FSteps[7].Children[1].Result := E_Result.Error;
FSteps[7].Children[1].Ready := FALSE;
FSteps[7].Children[1].Complete := TRUE;
FSteps[7].ExpectedDiagnosticCount := 1;
FSteps[7].ExpectedReleasedEntries[1] := 1;
FSteps[7].ExpectedResult := E_Result.Error;
{endregion}

{region "08 - No additional diagnostic or dispatch in Idle"}
FSteps[8].Task := E_OrchestratorTask.Idle;
FSteps[8].Children[1].State := E_State.Completed;
FSteps[8].Children[1].Result := E_Result.Error;
FSteps[8].Children[1].Ready := FALSE;
FSteps[8].Children[1].Complete := TRUE;
FSteps[8].ExpectedDiagnosticCount := 1;
FSteps[8].ExpectedResult := E_Result.Error;
{endregion}
END_METHOD

END_FUNCTION_BLOCK

// ---- SelfTests/TestCases/TestSuite_Orchestrator/Test_OrchestratorRepeatAfterReset.TcPOU
{region 'Documentation'}
(*!
<summary>Runs all three children twice with intervening Reset and without reinitializing the subject or capture.</summary>
*)
{endregion}
FUNCTION_BLOCK Test_OrchestratorRepeatAfterReset EXTENDS OrchestrationTestBase

SUPER^();

{region 'Documentation'}
(*!
<summary>Defines independent stimuli and expected requests, reservations, task status and diagnostic counts.</summary>
*)
{endregion}
METHOD PROTECTED ConfigureScenario
FStepCount := 21;

{region "01 - Idle readiness before child processing"}
FSteps[1].Task := E_OrchestratorTask.Idle;
FSteps[1].ExpectedReady := TRUE;
{endregion}

{region "02 - First child completes on its Start call"}
FSteps[2].Children[1].State := E_State.Completed;
FSteps[2].Children[1].Result := E_Result.Passed;
FSteps[2].Children[1].Ready := FALSE;
FSteps[2].Children[1].Complete := TRUE;
FSteps[2].ExpectedStartChild := 1;
FSteps[2].ExpectedSlot := 1;
FSteps[2].ExpectedReservations[1] := 1;
{endregion}

{region "03 - Observe first completion"}
FSteps[3].Children[1].State := E_State.Completed;
FSteps[3].Children[1].Result := E_Result.Passed;
FSteps[3].Children[1].Ready := FALSE;
FSteps[3].Children[1].Complete := TRUE;
FSteps[3].ExpectedSlot := 2;
FSteps[3].ExpectedReleasedEntries[1] := 1;
{endregion}

{region "04 - Second child completes on its Start call"}
FSteps[4].Children[1].State := E_State.Completed;
FSteps[4].Children[1].Result := E_Result.Passed;
FSteps[4].Children[1].Ready := FALSE;
FSteps[4].Children[1].Complete := TRUE;
FSteps[4].Children[2].State := E_State.Completed;
FSteps[4].Children[2].Result := E_Result.Passed;
FSteps[4].Children[2].Ready := FALSE;
FSteps[4].Children[2].Complete := TRUE;
FSteps[4].ExpectedStartChild := 2;
FSteps[4].ExpectedSlot := 2;
FSteps[4].ExpectedReservations[2] := 1;
{endregion}

{region "05 - Observe second completion"}
FSteps[5].Children[1].State := E_State.Completed;
FSteps[5].Children[1].Result := E_Result.Passed;
FSteps[5].Children[1].Ready := FALSE;
FSteps[5].Children[1].Complete := TRUE;
FSteps[5].Children[2].State := E_State.Completed;
FSteps[5].Children[2].Result := E_Result.Passed;
FSteps[5].Children[2].Ready := FALSE;
FSteps[5].Children[2].Complete := TRUE;
FSteps[5].ExpectedSlot := 3;
FSteps[5].ExpectedReleasedEntries[2] := 1;
{endregion}

{region "06 - Third child completes on its Start call"}
FSteps[6].Children[1].State := E_State.Completed;
FSteps[6].Children[1].Result := E_Result.Passed;
FSteps[6].Children[1].Ready := FALSE;
FSteps[6].Children[1].Complete := TRUE;
FSteps[6].Children[2].State := E_State.Completed;
FSteps[6].Children[2].Result := E_Result.Passed;
FSteps[6].Children[2].Ready := FALSE;
FSteps[6].Children[2].Complete := TRUE;
FSteps[6].Children[3].State := E_State.Completed;
FSteps[6].Children[3].Result := E_Result.Passed;
FSteps[6].Children[3].Ready := FALSE;
FSteps[6].Children[3].Complete := TRUE;
FSteps[6].ExpectedStartChild := 3;
FSteps[6].ExpectedSlot := 3;
FSteps[6].ExpectedReservations[3] := 1;
{endregion}

{region "07 - Observe execution completion"}
FSteps[7].Children[1].State := E_State.Completed;
FSteps[7].Children[1].Result := E_Result.Passed;
FSteps[7].Children[1].Ready := FALSE;
FSteps[7].Children[1].Complete := TRUE;
FSteps[7].Children[2].State := E_State.Completed;
FSteps[7].Children[2].Result := E_Result.Passed;
FSteps[7].Children[2].Ready := FALSE;
FSteps[7].Children[2].Complete := TRUE;
FSteps[7].Children[3].State := E_State.Completed;
FSteps[7].Children[3].Result := E_Result.Passed;
FSteps[7].Children[3].Ready := FALSE;
FSteps[7].Children[3].Complete := TRUE;
FSteps[7].ExpectedReleasedEntries[3] := 1;
FSteps[7].ExpectedFinished := TRUE;
{endregion}

{region "08 - Completed Execution task is retained"}
FSteps[8].Children[1].State := E_State.Completed;
FSteps[8].Children[1].Result := E_Result.Passed;
FSteps[8].Children[1].Ready := FALSE;
FSteps[8].Children[1].Complete := TRUE;
FSteps[8].Children[2].State := E_State.Completed;
FSteps[8].Children[2].Result := E_Result.Passed;
FSteps[8].Children[2].Ready := FALSE;
FSteps[8].Children[2].Complete := TRUE;
FSteps[8].Children[3].State := E_State.Completed;
FSteps[8].Children[3].Result := E_Result.Passed;
FSteps[8].Children[3].Ready := FALSE;
FSteps[8].Children[3].Complete := TRUE;
FSteps[8].ExpectedFinished := TRUE;
{endregion}

{region "09 - Reset first completed child"}
FSteps[9].Task := E_OrchestratorTask.Reset;
FSteps[9].Children[2].State := E_State.Completed;
FSteps[9].Children[2].Result := E_Result.Passed;
FSteps[9].Children[2].Ready := FALSE;
FSteps[9].Children[2].Complete := TRUE;
FSteps[9].Children[3].State := E_State.Completed;
FSteps[9].Children[3].Result := E_Result.Passed;
FSteps[9].Children[3].Ready := FALSE;
FSteps[9].Children[3].Complete := TRUE;
FSteps[9].ExpectedResetChild := 1;
FSteps[9].ExpectedReservations[1] := 1;
{endregion}

{region "10 - Release first and Reset second"}
FSteps[10].Task := E_OrchestratorTask.Reset;
FSteps[10].Children[3].State := E_State.Completed;
FSteps[10].Children[3].Result := E_Result.Passed;
FSteps[10].Children[3].Ready := FALSE;
FSteps[10].Children[3].Complete := TRUE;
FSteps[10].ExpectedResetChild := 2;
FSteps[10].ExpectedReservations[2] := 1;
FSteps[10].ExpectedReleasedEntries[1] := 1;
{endregion}

{region "11 - Release second and Reset third"}
FSteps[11].Task := E_OrchestratorTask.Reset;
FSteps[11].ExpectedResetChild := 3;
FSteps[11].ExpectedReservations[3] := 1;
FSteps[11].ExpectedReleasedEntries[2] := 1;
{endregion}

{region "12 - Observe full Reset completion"}
FSteps[12].Task := E_OrchestratorTask.Reset;
FSteps[12].ExpectedReleasedEntries[3] := 1;
FSteps[12].ExpectedResetFinished := TRUE;
{endregion}

{region "13 - Holding Reset must not reissue requests"}
FSteps[13].Task := E_OrchestratorTask.Reset;
FSteps[13].ExpectedResetFinished := TRUE;
{endregion}

{region "14 - Return to ready Idle"}
FSteps[14].Task := E_OrchestratorTask.Idle;
FSteps[14].ExpectedReady := TRUE;
{endregion}

{region "15 - First child completes on its Start call"}
FSteps[15].Children[1].State := E_State.Completed;
FSteps[15].Children[1].Result := E_Result.Passed;
FSteps[15].Children[1].Ready := FALSE;
FSteps[15].Children[1].Complete := TRUE;
FSteps[15].ExpectedStartChild := 1;
FSteps[15].ExpectedSlot := 1;
FSteps[15].ExpectedReservations[1] := 1;
{endregion}

{region "16 - Observe first completion"}
FSteps[16].Children[1].State := E_State.Completed;
FSteps[16].Children[1].Result := E_Result.Passed;
FSteps[16].Children[1].Ready := FALSE;
FSteps[16].Children[1].Complete := TRUE;
FSteps[16].ExpectedSlot := 2;
FSteps[16].ExpectedReleasedEntries[1] := 1;
{endregion}

{region "17 - Second child completes on its Start call"}
FSteps[17].Children[1].State := E_State.Completed;
FSteps[17].Children[1].Result := E_Result.Passed;
FSteps[17].Children[1].Ready := FALSE;
FSteps[17].Children[1].Complete := TRUE;
FSteps[17].Children[2].State := E_State.Completed;
FSteps[17].Children[2].Result := E_Result.Passed;
FSteps[17].Children[2].Ready := FALSE;
FSteps[17].Children[2].Complete := TRUE;
FSteps[17].ExpectedStartChild := 2;
FSteps[17].ExpectedSlot := 2;
FSteps[17].ExpectedReservations[2] := 1;
{endregion}

{region "18 - Observe second completion"}
FSteps[18].Children[1].State := E_State.Completed;
FSteps[18].Children[1].Result := E_Result.Passed;
FSteps[18].Children[1].Ready := FALSE;
FSteps[18].Children[1].Complete := TRUE;
FSteps[18].Children[2].State := E_State.Completed;
FSteps[18].Children[2].Result := E_Result.Passed;
FSteps[18].Children[2].Ready := FALSE;
FSteps[18].Children[2].Complete := TRUE;
FSteps[18].ExpectedSlot := 3;
FSteps[18].ExpectedReleasedEntries[2] := 1;
{endregion}

{region "19 - Third child completes on its Start call"}
FSteps[19].Children[1].State := E_State.Completed;
FSteps[19].Children[1].Result := E_Result.Passed;
FSteps[19].Children[1].Ready := FALSE;
FSteps[19].Children[1].Complete := TRUE;
FSteps[19].Children[2].State := E_State.Completed;
FSteps[19].Children[2].Result := E_Result.Passed;
FSteps[19].Children[2].Ready := FALSE;
FSteps[19].Children[2].Complete := TRUE;
FSteps[19].Children[3].State := E_State.Completed;
FSteps[19].Children[3].Result := E_Result.Passed;
FSteps[19].Children[3].Ready := FALSE;
FSteps[19].Children[3].Complete := TRUE;
FSteps[19].ExpectedStartChild := 3;
FSteps[19].ExpectedSlot := 3;
FSteps[19].ExpectedReservations[3] := 1;
{endregion}

{region "20 - Observe execution completion"}
FSteps[20].Children[1].State := E_State.Completed;
FSteps[20].Children[1].Result := E_Result.Passed;
FSteps[20].Children[1].Ready := FALSE;
FSteps[20].Children[1].Complete := TRUE;
FSteps[20].Children[2].State := E_State.Completed;
FSteps[20].Children[2].Result := E_Result.Passed;
FSteps[20].Children[2].Ready := FALSE;
FSteps[20].Children[2].Complete := TRUE;
FSteps[20].Children[3].State := E_State.Completed;
FSteps[20].Children[3].Result := E_Result.Passed;
FSteps[20].Children[3].Ready := FALSE;
FSteps[20].Children[3].Complete := TRUE;
FSteps[20].ExpectedReleasedEntries[3] := 1;
FSteps[20].ExpectedFinished := TRUE;
{endregion}

{region "21 - Completed Execution task is retained"}
FSteps[21].Children[1].State := E_State.Completed;
FSteps[21].Children[1].Result := E_Result.Passed;
FSteps[21].Children[1].Ready := FALSE;
FSteps[21].Children[1].Complete := TRUE;
FSteps[21].Children[2].State := E_State.Completed;
FSteps[21].Children[2].Result := E_Result.Passed;
FSteps[21].Children[2].Ready := FALSE;
FSteps[21].Children[2].Complete := TRUE;
FSteps[21].Children[3].State := E_State.Completed;
FSteps[21].Children[3].Result := E_Result.Passed;
FSteps[21].Children[3].Ready := FALSE;
FSteps[21].Children[3].Complete := TRUE;
FSteps[21].ExpectedFinished := TRUE;
{endregion}
END_METHOD

END_FUNCTION_BLOCK

// ---- SelfTests/TestCases/TestSuite_Orchestrator/Test_OrchestratorExecutionCapacityWait.TcPOU
{region 'Documentation'}
(*!
<summary>Waits silently for execution capacity, then starts each child exactly once without skipping the waiting candidate.</summary>
<description>
A ready first child cannot reserve for three calls, as with a slow event consumer.
Reservation responses apply before the helper; child state responses apply afterwards.
The second child proves correct continuation after capacity returns.
</description>
*)
{endregion}
FUNCTION_BLOCK Test_OrchestratorExecutionCapacityWait EXTENDS OrchestrationTestBase

SUPER^();

{region 'Documentation'}
(*!
<summary>Defines reservation responses and independent per-cycle expectations.</summary>
*)
{endregion}
METHOD PROTECTED ConfigureScenario
FChildCount := 2;
FStepCount := 10;

{region "01 - Observe initial readiness"}
FSteps[1].Task := E_OrchestratorTask.Idle;
FSteps[1].ExpectedReady := TRUE;
{endregion}

{region "02 - Wait for first child execution capacity"}
FSteps[2].ExecutionReservationResults[1] := E_EventReservationResult.WaitingForCapacity;
FSteps[2].ExpectedUnacceptedExecutionReservations[1] := 1;
FSteps[2].ExpectedSlot := 1;
{endregion}

{region "03 - Wait for first child execution capacity"}
FSteps[3].ExecutionReservationResults[1] := E_EventReservationResult.WaitingForCapacity;
FSteps[3].ExpectedUnacceptedExecutionReservations[1] := 1;
FSteps[3].ExpectedSlot := 1;
{endregion}

{region "04 - Wait for first child execution capacity"}
FSteps[4].ExecutionReservationResults[1] := E_EventReservationResult.WaitingForCapacity;
FSteps[4].ExpectedUnacceptedExecutionReservations[1] := 1;
FSteps[4].ExpectedSlot := 1;
{endregion}

{region "05 - Capacity restored - start first child"}
FSteps[5].Children[1].State := E_State.Running;
FSteps[5].Children[1].Ready := FALSE;
FSteps[5].ExpectedStartChild := 1;
FSteps[5].ExpectedSlot := 1;
FSteps[5].ExpectedReservations[1] := 1;
{endregion}

{region "06 - First child completes without another Start"}
FSteps[6].Children[1].State := E_State.Completed;
FSteps[6].Children[1].Ready := FALSE;
FSteps[6].Children[1].Complete := TRUE;
FSteps[6].Children[1].Result := E_Result.Passed;
FSteps[6].ExpectedSlot := 1;
FSteps[6].ExpectedReservations[1] := 1;
{endregion}

{region "07 - Release first child and select successor"}
FSteps[7].Children[1].State := E_State.Completed;
FSteps[7].Children[1].Ready := FALSE;
FSteps[7].Children[1].Complete := TRUE;
FSteps[7].Children[1].Result := E_Result.Passed;
FSteps[7].ExpectedSlot := 2;
FSteps[7].ExpectedReleasedEntries[1] := 1;
{endregion}

{region "08 - Start second child exactly once"}
FSteps[8].Children[1].State := E_State.Completed;
FSteps[8].Children[1].Ready := FALSE;
FSteps[8].Children[1].Complete := TRUE;
FSteps[8].Children[1].Result := E_Result.Passed;
FSteps[8].Children[2].State := E_State.Completed;
FSteps[8].Children[2].Ready := FALSE;
FSteps[8].Children[2].Complete := TRUE;
FSteps[8].Children[2].Result := E_Result.Passed;
FSteps[8].ExpectedStartChild := 2;
FSteps[8].ExpectedSlot := 2;
FSteps[8].ExpectedReservations[2] := 1;
{endregion}

{region "09 - Release second child and finish"}
FSteps[9].Children[1].State := E_State.Completed;
FSteps[9].Children[1].Ready := FALSE;
FSteps[9].Children[1].Complete := TRUE;
FSteps[9].Children[1].Result := E_Result.Passed;
FSteps[9].Children[2].State := E_State.Completed;
FSteps[9].Children[2].Ready := FALSE;
FSteps[9].Children[2].Complete := TRUE;
FSteps[9].Children[2].Result := E_Result.Passed;
FSteps[9].ExpectedFinished := TRUE;
FSteps[9].ExpectedReleasedEntries[2] := 1;
{endregion}

{region "10 - Completion remains stable without redispatch"}
FSteps[10].Children[1].State := E_State.Completed;
FSteps[10].Children[1].Ready := FALSE;
FSteps[10].Children[1].Complete := TRUE;
FSteps[10].Children[1].Result := E_Result.Passed;
FSteps[10].Children[2].State := E_State.Completed;
FSteps[10].Children[2].Ready := FALSE;
FSteps[10].Children[2].Complete := TRUE;
FSteps[10].Children[2].Result := E_Result.Passed;
FSteps[10].ExpectedFinished := TRUE;
{endregion}
END_METHOD

END_FUNCTION_BLOCK

// ---- SelfTests/TestCases/TestSuite_Orchestrator/Test_OrchestratorResetCapacityWait.TcPOU
{region 'Documentation'}
(*!
<summary>Retains Reset progress while capacity is unavailable, then resets the waiting child and its successor once.</summary>
<description>
Both children begin Completed. The first Reset reservation waits for three calls.
The subsequent Reset responses and releases prove no skipped child or duplicate request.
The final Idle call verifies that successful Reset restores readiness.
</description>
*)
{endregion}
FUNCTION_BLOCK Test_OrchestratorResetCapacityWait EXTENDS OrchestrationTestBase

SUPER^();

{region 'Documentation'}
(*!
<summary>Defines reservation responses and independent per-cycle expectations.</summary>
*)
{endregion}
METHOD PROTECTED ConfigureScenario
FChildCount := 2;
FStepCount := 10;

{region "01 - Establish terminal child observations"}
FSteps[1].Task := E_OrchestratorTask.Idle;
FSteps[1].Children[1].State := E_State.Completed;
FSteps[1].Children[1].Ready := FALSE;
FSteps[1].Children[1].Complete := TRUE;
FSteps[1].Children[1].Result := E_Result.Passed;
FSteps[1].Children[2].State := E_State.Completed;
FSteps[1].Children[2].Ready := FALSE;
FSteps[1].Children[2].Complete := TRUE;
FSteps[1].Children[2].Result := E_Result.Passed;
FSteps[1].ExpectedReady := TRUE;
{endregion}

{region "02 - Wait at first child without skipping to second"}
FSteps[2].Task := E_OrchestratorTask.Reset;
FSteps[2].Children[1].State := E_State.Completed;
FSteps[2].Children[1].Ready := FALSE;
FSteps[2].Children[1].Complete := TRUE;
FSteps[2].Children[1].Result := E_Result.Passed;
FSteps[2].Children[2].State := E_State.Completed;
FSteps[2].Children[2].Ready := FALSE;
FSteps[2].Children[2].Complete := TRUE;
FSteps[2].Children[2].Result := E_Result.Passed;
FSteps[2].ResetReservationResults[1] := E_EventReservationResult.WaitingForCapacity;
FSteps[2].ExpectedUnacceptedResetReservations[1] := 1;
{endregion}

{region "03 - Wait at first child without skipping to second"}
FSteps[3].Task := E_OrchestratorTask.Reset;
FSteps[3].Children[1].State := E_State.Completed;
FSteps[3].Children[1].Ready := FALSE;
FSteps[3].Children[1].Complete := TRUE;
FSteps[3].Children[1].Result := E_Result.Passed;
FSteps[3].Children[2].State := E_State.Completed;
FSteps[3].Children[2].Ready := FALSE;
FSteps[3].Children[2].Complete := TRUE;
FSteps[3].Children[2].Result := E_Result.Passed;
FSteps[3].ResetReservationResults[1] := E_EventReservationResult.WaitingForCapacity;
FSteps[3].ExpectedUnacceptedResetReservations[1] := 1;
{endregion}

{region "04 - Wait at first child without skipping to second"}
FSteps[4].Task := E_OrchestratorTask.Reset;
FSteps[4].Children[1].State := E_State.Completed;
FSteps[4].Children[1].Ready := FALSE;
FSteps[4].Children[1].Complete := TRUE;
FSteps[4].Children[1].Result := E_Result.Passed;
FSteps[4].Children[2].State := E_State.Completed;
FSteps[4].Children[2].Ready := FALSE;
FSteps[4].Children[2].Complete := TRUE;
FSteps[4].Children[2].Result := E_Result.Passed;
FSteps[4].ResetReservationResults[1] := E_EventReservationResult.WaitingForCapacity;
FSteps[4].ExpectedUnacceptedResetReservations[1] := 1;
{endregion}

{region "05 - Capacity restored - reset first child"}
FSteps[5].Task := E_OrchestratorTask.Reset;
FSteps[5].Children[1].State := E_State.Reset;
FSteps[5].Children[1].Ready := FALSE;
FSteps[5].Children[2].State := E_State.Completed;
FSteps[5].Children[2].Ready := FALSE;
FSteps[5].Children[2].Complete := TRUE;
FSteps[5].Children[2].Result := E_Result.Passed;
FSteps[5].ExpectedResetChild := 1;
FSteps[5].ExpectedReservations[1] := 1;
{endregion}

{region "06 - Reset second child while first reaches Idle"}
FSteps[6].Task := E_OrchestratorTask.Reset;
FSteps[6].Children[2].State := E_State.Reset;
FSteps[6].Children[2].Ready := FALSE;
FSteps[6].ExpectedResetChild := 2;
FSteps[6].ExpectedReservations[1] := 1;
FSteps[6].ExpectedReservations[2] := 1;
{endregion}

{region "07 - Release first child while second reaches Idle"}
FSteps[7].Task := E_OrchestratorTask.Reset;
FSteps[7].ExpectedReleasedEntries[1] := 1;
FSteps[7].ExpectedReservations[2] := 1;
{endregion}

{region "08 - Release second child and observe Reset completion"}
FSteps[8].Task := E_OrchestratorTask.Reset;
FSteps[8].ExpectedReleasedEntries[2] := 1;
FSteps[8].ExpectedResetFinished := TRUE;
{endregion}

{region "09 - No duplicate Reset after completion"}
FSteps[9].Task := E_OrchestratorTask.Reset;
FSteps[9].ExpectedResetFinished := TRUE;
{endregion}

{region "10 - Return to ready Idle with no remaining reservations"}
FSteps[10].Task := E_OrchestratorTask.Idle;
FSteps[10].ExpectedReady := TRUE;
{endregion}
END_METHOD

END_FUNCTION_BLOCK

// ---- SelfTests/TestCases/TestSuite_Orchestrator/Test_OrchestratorExecutionBudgetError.TcPOU
{region 'Documentation'}
(*!
<summary>Rejects an impossible execution budget without Start, capacity retry or repeated diagnostics.</summary>
<description>
The child returns Error, representing a budget larger than the configured buffer can hold.
Repeated Execution calls verify held Error and one diagnostic without further admission attempts.
Actual budget arithmetic belongs to reservation integration tests.
</description>
*)
{endregion}
FUNCTION_BLOCK Test_OrchestratorExecutionBudgetError EXTENDS OrchestrationTestBase

SUPER^();

{region 'Documentation'}
(*!
<summary>Defines reservation responses and independent per-cycle expectations.</summary>
*)
{endregion}
METHOD PROTECTED ConfigureScenario
FChildCount := 2;
FStepCount := 5;

{region "01 - Observe readiness before execution admission"}
FSteps[1].Task := E_OrchestratorTask.Idle;
FSteps[1].ExpectedReady := TRUE;
{endregion}

{region "02 - Reject the impossible execution reservation"}
FSteps[2].ExecutionReservationResults[1] := E_EventReservationResult.Error;
FSteps[2].ExpectedUnacceptedExecutionReservations[1] := 1;
FSteps[2].ExpectedSlot := 1;
FSteps[2].ExpectedResult := E_Result.Error;
FSteps[2].ExpectedDiagnosticCount := 1;
{endregion}

{region "03 - Retain Error without retry or another diagnostic"}
FSteps[3].ExecutionReservationResults[1] := E_EventReservationResult.Error;
FSteps[3].ExpectedSlot := 1;
FSteps[3].ExpectedResult := E_Result.Error;
FSteps[3].ExpectedDiagnosticCount := 1;
{endregion}

{region "04 - Retain Error without retry or another diagnostic"}
FSteps[4].ExecutionReservationResults[1] := E_EventReservationResult.Error;
FSteps[4].ExpectedSlot := 1;
FSteps[4].ExpectedResult := E_Result.Error;
FSteps[4].ExpectedDiagnosticCount := 1;
{endregion}

{region "05 - Retain Error without retry or another diagnostic"}
FSteps[5].ExecutionReservationResults[1] := E_EventReservationResult.Error;
FSteps[5].ExpectedSlot := 1;
FSteps[5].ExpectedResult := E_Result.Error;
FSteps[5].ExpectedDiagnosticCount := 1;
{endregion}
END_METHOD

END_FUNCTION_BLOCK

// ---- SelfTests/TestSuites/TestSuite_SerialOrchestration.TcPOU
{region 'Documentation'}
(*!
<summary>Verifies Serial-specific registration order, admission and child progression.</summary>
*)
{endregion}
FUNCTION_BLOCK TestSuite_SerialOrchestration EXTENDS TestSuiteBase
VAR
    FRegistrationOrder : Test_SerialRegistrationOrder;
    FImmediateCompletion : Test_SerialImmediateCompletion;
    FUnequalDurations : Test_SerialUnequalDurations;
    FNotReadyCandidate : Test_SerialNotReadyCandidate;
    FFailedResultContinues : Test_SerialFailedResultContinues;
    FTestCases : ARRAY[1..TestCaseCapacity] OF I_TestCase;
END_VAR
VAR CONSTANT
    TestCaseCapacity : UINT := 5;
END_VAR

SUPER^();

{region 'Documentation'}
(*!
<summary>Initializes and registers the owned orchestration scenarios in deterministic order.</summary>
*)
{endregion}
METHOD PROTECTED Configure
VAR_IN_OUT
    // SA0167: Borrowed builder; VAR_IN_OUT creates no temporary instance.
    {attribute 'analysis' := '-167'}
    Builder : TestSuiteConfigurationBuilder; //! Borrowed owner configuration builder used only during this Configure call; register this owner's concrete children.
END_VAR
VAR
    TestConfig : ST_TestCaseConfig;
END_VAR
Builder.Initialize(Mode := E_OrchestrationMode.Serial,
    TestCases := FTestCases);

FRegistrationOrder.Initialize(Parent := THIS^,
    TestName := 'RegistrationOrder',
    Config := TestConfig);
Builder.Register(TestCase := FRegistrationOrder);

FImmediateCompletion.Initialize(Parent := THIS^,
    TestName := 'ImmediateCompletion',
    Config := TestConfig);
Builder.Register(TestCase := FImmediateCompletion);

FUnequalDurations.Initialize(Parent := THIS^,
    TestName := 'UnequalDurations',
    Config := TestConfig);
Builder.Register(TestCase := FUnequalDurations);

FNotReadyCandidate.Initialize(Parent := THIS^,
    TestName := 'NotReadyCandidate',
    Config := TestConfig);
Builder.Register(TestCase := FNotReadyCandidate);

FFailedResultContinues.Initialize(Parent := THIS^,
    TestName := 'FailedResultContinues',
    Config := TestConfig);
Builder.Register(TestCase := FFailedResultContinues);
END_METHOD

{region 'Documentation'}
(*!
<summary>Returns the registered Test Case from the same array used during configuration.</summary>
*)
{endregion}
METHOD PUBLIC GetTestCase : I_TestCase //! Typed child interface at the original array index; zero when no entry is available.
VAR_INPUT
    Index : DINT; //! Original occupied child-array index, rather than an ordinal position.
END_VAR
GetTestCase := 0;
IF (ChildCount = 0) OR (Index < ChildArrayLowerBound)
    OR (DINT_TO_LINT(Index) >= DINT_TO_LINT(ChildArrayLowerBound) + UINT_TO_LINT(ChildCount)) THEN
    RETURN;
END_IF;

GetTestCase := FTestCases[Index];
END_METHOD

{region 'Documentation'}
(*!
<summary>Calls each owned Test Case once per initialized Suite cycle, including completion.</summary>
*)
{endregion}
METHOD PROTECTED ProcessTestCases
FRegistrationOrder();
FImmediateCompletion();
FUnequalDurations();
FNotReadyCandidate();
FFailedResultContinues();
END_METHOD

END_FUNCTION_BLOCK

// ---- SelfTests/TestCases/TestSuite_SerialOrchestration/Test_SerialRegistrationOrder.TcPOU
{region 'Documentation'}
(*!
<summary>Checks A-B-C registration order, delayed observation and exactly one active child.</summary>
*)
{endregion}
FUNCTION_BLOCK Test_SerialRegistrationOrder EXTENDS OrchestrationTestBase

SUPER^();

{region 'Documentation'}
(*!
<summary>Defines this scenario independently of the subject's internal fields.</summary>
*)
{endregion}
METHOD PROTECTED ConfigureScenario
FArrayLayout := E_OrchestrationArrayLayout.Ordinary;
FChildCount := 3;
ConfigureStandardSequence();
END_METHOD

END_FUNCTION_BLOCK

// ---- SelfTests/TestCases/TestSuite_SerialOrchestration/Test_SerialImmediateCompletion.TcPOU
{region 'Documentation'}
(*!
<summary>Checks children already Completed at the first helper call after their Start.</summary>
*)
{endregion}
FUNCTION_BLOCK Test_SerialImmediateCompletion EXTENDS OrchestrationTestBase

SUPER^();

{region 'Documentation'}
(*!
<summary>Defines this scenario independently of the subject's internal fields.</summary>
*)
{endregion}
METHOD PROTECTED ConfigureScenario
FArrayLayout := E_OrchestrationArrayLayout.Ordinary;
FChildCount := 3;
FStepCount := 8;

{region "Cycle 01 - Idle readiness"}
FSteps[1].Task := E_OrchestratorTask.Idle;
FSteps[1].ExpectedReady := TRUE;
{endregion}

{region "Cycle 02 - Start child 1"}
FSteps[2].Children[1].State := E_State.Completed;
FSteps[2].Children[1].Ready := FALSE;
FSteps[2].Children[1].Complete := TRUE;
FSteps[2].Children[1].Result := E_Result.Passed;
FSteps[2].ExpectedStartChild := 1;
FSteps[2].ExpectedSlot := 1;
FSteps[2].ExpectedReservations[1] := 1;
{endregion}

{region "Cycle 03 - Reconcile completed child 1"}
FSteps[3].Children[1].State := E_State.Completed;
FSteps[3].Children[1].Ready := FALSE;
FSteps[3].Children[1].Complete := TRUE;
FSteps[3].Children[1].Result := E_Result.Passed;
FSteps[3].ExpectedSlot := 2;
FSteps[3].ExpectedReleasedEntries[1] := 1;
{endregion}

{region "Cycle 04 - Start child 2"}
FSteps[4].Children[1].State := E_State.Completed;
FSteps[4].Children[1].Ready := FALSE;
FSteps[4].Children[1].Complete := TRUE;
FSteps[4].Children[1].Result := E_Result.Passed;
FSteps[4].Children[2].State := E_State.Completed;
FSteps[4].Children[2].Ready := FALSE;
FSteps[4].Children[2].Complete := TRUE;
FSteps[4].Children[2].Result := E_Result.Passed;
FSteps[4].ExpectedStartChild := 2;
FSteps[4].ExpectedSlot := 2;
FSteps[4].ExpectedReservations[2] := 1;
{endregion}

{region "Cycle 05 - Reconcile completed child 2"}
FSteps[5].Children[1].State := E_State.Completed;
FSteps[5].Children[1].Ready := FALSE;
FSteps[5].Children[1].Complete := TRUE;
FSteps[5].Children[1].Result := E_Result.Passed;
FSteps[5].Children[2].State := E_State.Completed;
FSteps[5].Children[2].Ready := FALSE;
FSteps[5].Children[2].Complete := TRUE;
FSteps[5].Children[2].Result := E_Result.Passed;
FSteps[5].ExpectedSlot := 3;
FSteps[5].ExpectedReleasedEntries[2] := 1;
{endregion}

{region "Cycle 06 - Start child 3"}
FSteps[6].Children[1].State := E_State.Completed;
FSteps[6].Children[1].Ready := FALSE;
FSteps[6].Children[1].Complete := TRUE;
FSteps[6].Children[1].Result := E_Result.Passed;
FSteps[6].Children[2].State := E_State.Completed;
FSteps[6].Children[2].Ready := FALSE;
FSteps[6].Children[2].Complete := TRUE;
FSteps[6].Children[2].Result := E_Result.Passed;
FSteps[6].Children[3].State := E_State.Completed;
FSteps[6].Children[3].Ready := FALSE;
FSteps[6].Children[3].Complete := TRUE;
FSteps[6].Children[3].Result := E_Result.Passed;
FSteps[6].ExpectedStartChild := 3;
FSteps[6].ExpectedSlot := 3;
FSteps[6].ExpectedReservations[3] := 1;
{endregion}

{region "Cycle 07 - Completed observation"}
FSteps[7].Children[1].State := E_State.Completed;
FSteps[7].Children[1].Ready := FALSE;
FSteps[7].Children[1].Complete := TRUE;
FSteps[7].Children[1].Result := E_Result.Passed;
FSteps[7].Children[2].State := E_State.Completed;
FSteps[7].Children[2].Ready := FALSE;
FSteps[7].Children[2].Complete := TRUE;
FSteps[7].Children[2].Result := E_Result.Passed;
FSteps[7].Children[3].State := E_State.Completed;
FSteps[7].Children[3].Ready := FALSE;
FSteps[7].Children[3].Complete := TRUE;
FSteps[7].Children[3].Result := E_Result.Passed;
FSteps[7].ExpectedReleasedEntries[3] := 1;
FSteps[7].ExpectedFinished := TRUE;
{endregion}

{region "Cycle 08 - Completed observation"}
FSteps[8].Children[1].State := E_State.Completed;
FSteps[8].Children[1].Ready := FALSE;
FSteps[8].Children[1].Complete := TRUE;
FSteps[8].Children[1].Result := E_Result.Passed;
FSteps[8].Children[2].State := E_State.Completed;
FSteps[8].Children[2].Ready := FALSE;
FSteps[8].Children[2].Complete := TRUE;
FSteps[8].Children[2].Result := E_Result.Passed;
FSteps[8].Children[3].State := E_State.Completed;
FSteps[8].Children[3].Ready := FALSE;
FSteps[8].Children[3].Complete := TRUE;
FSteps[8].Children[3].Result := E_Result.Passed;
FSteps[8].ExpectedFinished := TRUE;
{endregion}
END_METHOD

END_FUNCTION_BLOCK

// ---- SelfTests/TestCases/TestSuite_SerialOrchestration/Test_SerialUnequalDurations.TcPOU
{region 'Documentation'}
(*!
<summary>Checks long, immediate and shorter children; Completing is not terminal completion.</summary>
*)
{endregion}
FUNCTION_BLOCK Test_SerialUnequalDurations EXTENDS OrchestrationTestBase

SUPER^();

{region 'Documentation'}
(*!
<summary>Defines this scenario independently of the subject's internal fields.</summary>
*)
{endregion}
METHOD PROTECTED ConfigureScenario
FArrayLayout := E_OrchestrationArrayLayout.Ordinary;
FChildCount := 3;
FStepCount := 15;

{region "Cycle 01 - Idle readiness"}
FSteps[1].Task := E_OrchestratorTask.Idle;
FSteps[1].ExpectedReady := TRUE;
{endregion}

{region "Cycle 02 - Start child 1"}
FSteps[2].Children[1].State := E_State.Running;
FSteps[2].Children[1].Ready := FALSE;
FSteps[2].ExpectedStartChild := 1;
FSteps[2].ExpectedSlot := 1;
FSteps[2].ExpectedReservations[1] := 1;
{endregion}

{region "Cycle 03 - Child progress"}
FSteps[3].Children[1].State := E_State.Running;
FSteps[3].Children[1].Ready := FALSE;
FSteps[3].ExpectedSlot := 1;
FSteps[3].ExpectedReservations[1] := 1;
{endregion}

{region "Cycle 04 - Child progress"}
FSteps[4].Children[1].State := E_State.Running;
FSteps[4].Children[1].Ready := FALSE;
FSteps[4].ExpectedSlot := 1;
FSteps[4].ExpectedReservations[1] := 1;
{endregion}

{region "Cycle 05 - Child progress"}
FSteps[5].Children[1].State := E_State.Running;
FSteps[5].Children[1].Ready := FALSE;
FSteps[5].ExpectedSlot := 1;
FSteps[5].ExpectedReservations[1] := 1;
{endregion}

{region "Cycle 06 - Child progress"}
FSteps[6].Children[1].State := E_State.Completing;
FSteps[6].Children[1].Ready := FALSE;
FSteps[6].ExpectedSlot := 1;
FSteps[6].ExpectedReservations[1] := 1;
{endregion}

{region "Cycle 07 - Child progress"}
FSteps[7].Children[1].State := E_State.Completed;
FSteps[7].Children[1].Ready := FALSE;
FSteps[7].Children[1].Complete := TRUE;
FSteps[7].Children[1].Result := E_Result.Passed;
FSteps[7].ExpectedSlot := 1;
FSteps[7].ExpectedReservations[1] := 1;
{endregion}

{region "Cycle 08 - Reconcile completed child 1"}
FSteps[8].Children[1].State := E_State.Completed;
FSteps[8].Children[1].Ready := FALSE;
FSteps[8].Children[1].Complete := TRUE;
FSteps[8].Children[1].Result := E_Result.Passed;
FSteps[8].ExpectedSlot := 2;
FSteps[8].ExpectedReleasedEntries[1] := 1;
{endregion}

{region "Cycle 09 - Start child 2"}
FSteps[9].Children[1].State := E_State.Completed;
FSteps[9].Children[1].Ready := FALSE;
FSteps[9].Children[1].Complete := TRUE;
FSteps[9].Children[1].Result := E_Result.Passed;
FSteps[9].Children[2].State := E_State.Completed;
FSteps[9].Children[2].Ready := FALSE;
FSteps[9].Children[2].Complete := TRUE;
FSteps[9].Children[2].Result := E_Result.Passed;
FSteps[9].ExpectedStartChild := 2;
FSteps[9].ExpectedSlot := 2;
FSteps[9].ExpectedReservations[2] := 1;
{endregion}

{region "Cycle 10 - Reconcile completed child 2"}
FSteps[10].Children[1].State := E_State.Completed;
FSteps[10].Children[1].Ready := FALSE;
FSteps[10].Children[1].Complete := TRUE;
FSteps[10].Children[1].Result := E_Result.Passed;
FSteps[10].Children[2].State := E_State.Completed;
FSteps[10].Children[2].Ready := FALSE;
FSteps[10].Children[2].Complete := TRUE;
FSteps[10].Children[2].Result := E_Result.Passed;
FSteps[10].ExpectedSlot := 3;
FSteps[10].ExpectedReleasedEntries[2] := 1;
{endregion}

{region "Cycle 11 - Start child 3"}
FSteps[11].Children[1].State := E_State.Completed;
FSteps[11].Children[1].Ready := FALSE;
FSteps[11].Children[1].Complete := TRUE;
FSteps[11].Children[1].Result := E_Result.Passed;
FSteps[11].Children[2].State := E_State.Completed;
FSteps[11].Children[2].Ready := FALSE;
FSteps[11].Children[2].Complete := TRUE;
FSteps[11].Children[2].Result := E_Result.Passed;
FSteps[11].Children[3].State := E_State.Running;
FSteps[11].Children[3].Ready := FALSE;
FSteps[11].ExpectedStartChild := 3;
FSteps[11].ExpectedSlot := 3;
FSteps[11].ExpectedReservations[3] := 1;
{endregion}

{region "Cycle 12 - Child progress"}
FSteps[12].Children[1].State := E_State.Completed;
FSteps[12].Children[1].Ready := FALSE;
FSteps[12].Children[1].Complete := TRUE;
FSteps[12].Children[1].Result := E_Result.Passed;
FSteps[12].Children[2].State := E_State.Completed;
FSteps[12].Children[2].Ready := FALSE;
FSteps[12].Children[2].Complete := TRUE;
FSteps[12].Children[2].Result := E_Result.Passed;
FSteps[12].Children[3].State := E_State.Running;
FSteps[12].Children[3].Ready := FALSE;
FSteps[12].ExpectedSlot := 3;
FSteps[12].ExpectedReservations[3] := 1;
{endregion}

{region "Cycle 13 - Child progress"}
FSteps[13].Children[1].State := E_State.Completed;
FSteps[13].Children[1].Ready := FALSE;
FSteps[13].Children[1].Complete := TRUE;
FSteps[13].Children[1].Result := E_Result.Passed;
FSteps[13].Children[2].State := E_State.Completed;
FSteps[13].Children[2].Ready := FALSE;
FSteps[13].Children[2].Complete := TRUE;
FSteps[13].Children[2].Result := E_Result.Passed;
FSteps[13].Children[3].State := E_State.Completed;
FSteps[13].Children[3].Ready := FALSE;
FSteps[13].Children[3].Complete := TRUE;
FSteps[13].Children[3].Result := E_Result.Passed;
FSteps[13].ExpectedSlot := 3;
FSteps[13].ExpectedReservations[3] := 1;
{endregion}

{region "Cycle 14 - Completed observation"}
FSteps[14].Children[1].State := E_State.Completed;
FSteps[14].Children[1].Ready := FALSE;
FSteps[14].Children[1].Complete := TRUE;
FSteps[14].Children[1].Result := E_Result.Passed;
FSteps[14].Children[2].State := E_State.Completed;
FSteps[14].Children[2].Ready := FALSE;
FSteps[14].Children[2].Complete := TRUE;
FSteps[14].Children[2].Result := E_Result.Passed;
FSteps[14].Children[3].State := E_State.Completed;
FSteps[14].Children[3].Ready := FALSE;
FSteps[14].Children[3].Complete := TRUE;
FSteps[14].Children[3].Result := E_Result.Passed;
FSteps[14].ExpectedReleasedEntries[3] := 1;
FSteps[14].ExpectedFinished := TRUE;
{endregion}

{region "Cycle 15 - Completed observation"}
FSteps[15].Children[1].State := E_State.Completed;
FSteps[15].Children[1].Ready := FALSE;
FSteps[15].Children[1].Complete := TRUE;
FSteps[15].Children[1].Result := E_Result.Passed;
FSteps[15].Children[2].State := E_State.Completed;
FSteps[15].Children[2].Ready := FALSE;
FSteps[15].Children[2].Complete := TRUE;
FSteps[15].Children[2].Result := E_Result.Passed;
FSteps[15].Children[3].State := E_State.Completed;
FSteps[15].Children[3].Ready := FALSE;
FSteps[15].Children[3].Complete := TRUE;
FSteps[15].Children[3].Result := E_Result.Passed;
FSteps[15].ExpectedFinished := TRUE;
{endregion}
END_METHOD

END_FUNCTION_BLOCK

// ---- SelfTests/TestCases/TestSuite_SerialOrchestration/Test_SerialNotReadyCandidate.TcPOU
{region 'Documentation'}
(*!
<summary>Rejects the next serial candidate when not ready; no reservation or later Start is permitted.</summary>
*)
{endregion}
FUNCTION_BLOCK Test_SerialNotReadyCandidate EXTENDS OrchestrationTestBase

SUPER^();

{region 'Documentation'}
(*!
<summary>Defines independent stimuli and expected requests, reservations, task status and diagnostic counts.</summary>
*)
{endregion}
METHOD PROTECTED ConfigureScenario
FStepCount := 7;

{region "01 - Idle readiness before child processing"}
FSteps[1].Task := E_OrchestratorTask.Idle;
FSteps[1].ExpectedReady := TRUE;
{endregion}

{region "02 - Start first child; next child loses readiness"}
FSteps[2].Children[1].State := E_State.Running;
FSteps[2].Children[1].Ready := FALSE;
FSteps[2].Children[2].Ready := FALSE;
FSteps[2].ExpectedStartChild := 1;
FSteps[2].ExpectedSlot := 1;
FSteps[2].ExpectedReservations[1] := 1;
{endregion}

{region "03 - First child completes; next remains not ready"}
FSteps[3].Children[1].State := E_State.Completed;
FSteps[3].Children[1].Result := E_Result.Passed;
FSteps[3].Children[1].Ready := FALSE;
FSteps[3].Children[1].Complete := TRUE;
FSteps[3].Children[2].Ready := FALSE;
FSteps[3].ExpectedSlot := 1;
FSteps[3].ExpectedReservations[1] := 1;
{endregion}

{region "04 - Reconcile first child and select second slot"}
FSteps[4].Children[1].State := E_State.Completed;
FSteps[4].Children[1].Result := E_Result.Passed;
FSteps[4].Children[1].Ready := FALSE;
FSteps[4].Children[1].Complete := TRUE;
FSteps[4].Children[2].Ready := FALSE;
FSteps[4].ExpectedSlot := 2;
FSteps[4].ExpectedReleasedEntries[1] := 1;
{endregion}

{region "05 - Reject not-ready candidate"}
FSteps[5].Children[1].State := E_State.Completed;
FSteps[5].Children[1].Result := E_Result.Passed;
FSteps[5].Children[1].Ready := FALSE;
FSteps[5].Children[1].Complete := TRUE;
FSteps[5].Children[2].Ready := FALSE;
FSteps[5].ExpectedSlot := 2;
FSteps[5].ExpectedDiagnosticCount := 1;
FSteps[5].ExpectedResult := E_Result.Error;
{endregion}

{region "06 - Repeated failure does not publish again"}
FSteps[6].Children[1].State := E_State.Completed;
FSteps[6].Children[1].Result := E_Result.Passed;
FSteps[6].Children[1].Ready := FALSE;
FSteps[6].Children[1].Complete := TRUE;
FSteps[6].Children[2].Ready := FALSE;
FSteps[6].ExpectedSlot := 2;
FSteps[6].ExpectedDiagnosticCount := 1;
FSteps[6].ExpectedResult := E_Result.Error;
{endregion}

{region "07 - Idle stops dispatch but retains the error"}
FSteps[7].Task := E_OrchestratorTask.Idle;
FSteps[7].Children[1].State := E_State.Completed;
FSteps[7].Children[1].Result := E_Result.Passed;
FSteps[7].Children[1].Ready := FALSE;
FSteps[7].Children[1].Complete := TRUE;
FSteps[7].ExpectedDiagnosticCount := 1;
FSteps[7].ExpectedResult := E_Result.Error;
{endregion}
END_METHOD

END_FUNCTION_BLOCK

// ---- SelfTests/TestCases/TestSuite_SerialOrchestration/Test_SerialFailedResultContinues.TcPOU
{region 'Documentation'}
(*!
<summary>A normal Failed result does not become a helper Error or prevent later serial children.</summary>
*)
{endregion}
FUNCTION_BLOCK Test_SerialFailedResultContinues EXTENDS OrchestrationTestBase

SUPER^();

{region 'Documentation'}
(*!
<summary>Defines independent stimuli and expected requests, reservations, task status and diagnostic counts.</summary>
*)
{endregion}
METHOD PROTECTED ConfigureScenario
VAR
    Index : INT;
END_VAR
ConfigureStandardSequence();
// A completed Failed child remains a normal execution outcome, not a helper Error.
FOR Index := 4 TO FStepCount DO
    FSteps[Index].Children[1].Result := E_Result.Failed;
END_FOR;
END_METHOD

END_FUNCTION_BLOCK

// ---- SelfTests/TestSuites/TestSuite_ParallelOrchestration.TcPOU
{region 'Documentation'}
(*!
<summary>Runs focused Parallel Orchestrator scenarios serially with isolated child observations and diagnostics.</summary>
*)
{endregion}
FUNCTION_BLOCK TestSuite_ParallelOrchestration EXTENDS TestSuiteBase
VAR
    FUnequalDurations : Test_ParallelUnequalDurations;
    FFirstFittingAdmission : Test_ParallelFirstFittingAdmission;
    FMissingStartReaction : Test_ParallelMissingStartReaction;
    FReadinessLost : Test_ParallelReadinessLost;
    FFailedResultContinues : Test_ParallelFailedResultContinues;
    FChildError : Test_ParallelChildError;
    FAbortMixedProgress : Test_ParallelAbortMixedProgress;
    FResetOverlappingExecution : Test_ParallelResetOverlappingExecution;
    FTestCases : ARRAY[1..TestCaseCapacity] OF I_TestCase;
END_VAR
VAR CONSTANT
    TestCaseCapacity : UINT := 8;
END_VAR

SUPER^();

{region 'Documentation'}
(*!
<summary>Initializes and registers the owned orchestration scenarios in deterministic order.</summary>
*)
{endregion}
METHOD PROTECTED Configure
VAR_IN_OUT
    // SA0167: Borrowed builder; VAR_IN_OUT creates no temporary instance.
    {attribute 'analysis' := '-167'}
    Builder : TestSuiteConfigurationBuilder; //! Borrowed owner configuration builder used only during this Configure call; register this owner's concrete children.
END_VAR
VAR
    TestConfig : ST_TestCaseConfig;
END_VAR
Builder.Initialize(Mode := E_OrchestrationMode.Serial,
    TestCases := FTestCases);

FUnequalDurations.Initialize(Parent := THIS^,
    TestName := 'UnequalDurations',
    Config := TestConfig);
Builder.Register(TestCase := FUnequalDurations);

FFirstFittingAdmission.Initialize(Parent := THIS^,
    TestName := 'FirstFittingAdmission',
    Config := TestConfig);
Builder.Register(TestCase := FFirstFittingAdmission);

FMissingStartReaction.Initialize(Parent := THIS^,
    TestName := 'MissingStartReaction',
    Config := TestConfig);
Builder.Register(TestCase := FMissingStartReaction);

FReadinessLost.Initialize(Parent := THIS^,
    TestName := 'ReadinessLost',
    Config := TestConfig);
Builder.Register(TestCase := FReadinessLost);

FFailedResultContinues.Initialize(Parent := THIS^,
    TestName := 'FailedResultContinues',
    Config := TestConfig);
Builder.Register(TestCase := FFailedResultContinues);

FChildError.Initialize(Parent := THIS^,
    TestName := 'ChildError',
    Config := TestConfig);
Builder.Register(TestCase := FChildError);

FAbortMixedProgress.Initialize(Parent := THIS^,
    TestName := 'AbortMixedProgress',
    Config := TestConfig);
Builder.Register(TestCase := FAbortMixedProgress);

FResetOverlappingExecution.Initialize(Parent := THIS^,
    TestName := 'ResetOverlappingExecution',
    Config := TestConfig);
Builder.Register(TestCase := FResetOverlappingExecution);
END_METHOD

{region 'Documentation'}
(*!
<summary>Returns the registered Test Case from the same array used during configuration.</summary>
*)
{endregion}
METHOD PUBLIC GetTestCase : I_TestCase //! Typed child interface at the original array index; zero when no entry is available.
VAR_INPUT
    Index : DINT; //! Original occupied child-array index, rather than an ordinal position.
END_VAR
GetTestCase := 0;
IF (ChildCount = 0) OR (Index < ChildArrayLowerBound)
    OR (DINT_TO_LINT(Index) >= DINT_TO_LINT(ChildArrayLowerBound) + UINT_TO_LINT(ChildCount)) THEN
    RETURN;
END_IF;

GetTestCase := FTestCases[Index];
END_METHOD

{region 'Documentation'}
(*!
<summary>Calls each owned Test Case once per initialized Suite cycle, including completion.</summary>
*)
{endregion}
METHOD PROTECTED ProcessTestCases
FUnequalDurations();
FFirstFittingAdmission();
FMissingStartReaction();
FReadinessLost();
FFailedResultContinues();
FChildError();
FAbortMixedProgress();
FResetOverlappingExecution();
END_METHOD

END_FUNCTION_BLOCK

// ---- SelfTests/TestCases/TestSuite_ParallelOrchestration/Test_ParallelUnequalDurations.TcPOU
{region 'Documentation'}
(*!
<summary>Starts one same-slot child per cycle and waits for the last participant despite unequal and immediate completion.</summary>
<description>
Child 2 completes on its Start call while child 1 continues. Child 3 runs concurrently and
finishes before child 1. Completed children retain their terminal observations so
redispatch and premature group completion are detectable.
</description>
*)
{endregion}
FUNCTION_BLOCK Test_ParallelUnequalDurations EXTENDS OrchestrationTestBase

SUPER^();

{region 'Documentation'}
(*!
<summary>Defines independent per-cycle child responses and Parallel dispatch expectations.</summary>
*)
{endregion}
METHOD PROTECTED ConfigureScenario
FChildSlots[1] := 1;
FChildSlots[2] := 1;
FChildSlots[3] := 1;
FStepCount := 9;

{region "01 - Observe initial readiness"}
FSteps[1].Task := E_OrchestratorTask.Idle;
FSteps[1].ExpectedReady := TRUE;
{endregion}

{region "02 - Start long-running child 1"}
FSteps[2].Children[1].State := E_State.Running;
FSteps[2].Children[1].Ready := FALSE;
FSteps[2].ExpectedStartChild := 1;
FSteps[2].ExpectedSlot := 1;
FSteps[2].ExpectedReservations[1] := 1;
FSteps[2].MaxActiveChildCount := 1;
{endregion}

{region "03 - Start child 2 which completes immediately"}
FSteps[3].Children[1].State := E_State.Running;
FSteps[3].Children[1].Ready := FALSE;
FSteps[3].Children[2].State := E_State.Completed;
FSteps[3].Children[2].Ready := FALSE;
FSteps[3].Children[2].Complete := TRUE;
FSteps[3].Children[2].Result := E_Result.Passed;
FSteps[3].ExpectedStartChild := 2;
FSteps[3].ExpectedSlot := 1;
FSteps[3].ExpectedReservations[1] := 1;
FSteps[3].ExpectedReservations[2] := 1;
FSteps[3].MaxActiveChildCount := 2;
{endregion}

{region "04 - Release child 2 and start child 3 while child 1 runs"}
FSteps[4].Children[1].State := E_State.Running;
FSteps[4].Children[1].Ready := FALSE;
FSteps[4].Children[2].State := E_State.Completed;
FSteps[4].Children[2].Ready := FALSE;
FSteps[4].Children[2].Complete := TRUE;
FSteps[4].Children[2].Result := E_Result.Passed;
FSteps[4].Children[3].State := E_State.Running;
FSteps[4].Children[3].Ready := FALSE;
FSteps[4].ExpectedStartChild := 3;
FSteps[4].ExpectedSlot := 1;
FSteps[4].ExpectedReservations[1] := 1;
FSteps[4].ExpectedReservations[3] := 1;
FSteps[4].ExpectedReleasedEntries[2] := 1;
FSteps[4].MaxActiveChildCount := 2;
{endregion}

{region "05 - Keep children 1 and 3 running without redispatch"}
FSteps[5].Children[1].State := E_State.Running;
FSteps[5].Children[1].Ready := FALSE;
FSteps[5].Children[2].State := E_State.Completed;
FSteps[5].Children[2].Ready := FALSE;
FSteps[5].Children[2].Complete := TRUE;
FSteps[5].Children[2].Result := E_Result.Passed;
FSteps[5].Children[3].State := E_State.Running;
FSteps[5].Children[3].Ready := FALSE;
FSteps[5].ExpectedSlot := 1;
FSteps[5].ExpectedReservations[1] := 1;
FSteps[5].ExpectedReservations[3] := 1;
FSteps[5].MaxActiveChildCount := 2;
{endregion}

{region "06 - Child 3 completes while child 1 still runs"}
FSteps[6].Children[1].State := E_State.Running;
FSteps[6].Children[1].Ready := FALSE;
FSteps[6].Children[2].State := E_State.Completed;
FSteps[6].Children[2].Ready := FALSE;
FSteps[6].Children[2].Complete := TRUE;
FSteps[6].Children[2].Result := E_Result.Passed;
FSteps[6].Children[3].State := E_State.Completed;
FSteps[6].Children[3].Ready := FALSE;
FSteps[6].Children[3].Complete := TRUE;
FSteps[6].Children[3].Result := E_Result.Passed;
FSteps[6].ExpectedSlot := 1;
FSteps[6].ExpectedReservations[1] := 1;
FSteps[6].ExpectedReservations[3] := 1;
FSteps[6].MaxActiveChildCount := 2;
{endregion}

{region "07 - Release child 3 then observe child 1 completing"}
FSteps[7].Children[1].State := E_State.Completed;
FSteps[7].Children[1].Ready := FALSE;
FSteps[7].Children[1].Complete := TRUE;
FSteps[7].Children[1].Result := E_Result.Passed;
FSteps[7].Children[2].State := E_State.Completed;
FSteps[7].Children[2].Ready := FALSE;
FSteps[7].Children[2].Complete := TRUE;
FSteps[7].Children[2].Result := E_Result.Passed;
FSteps[7].Children[3].State := E_State.Completed;
FSteps[7].Children[3].Ready := FALSE;
FSteps[7].Children[3].Complete := TRUE;
FSteps[7].Children[3].Result := E_Result.Passed;
FSteps[7].ExpectedSlot := 1;
FSteps[7].ExpectedReservations[1] := 1;
FSteps[7].ExpectedReleasedEntries[3] := 1;
FSteps[7].MaxActiveChildCount := 1;
{endregion}

{region "08 - Reconcile the last reservation and finish the group"}
FSteps[8].Children[1].State := E_State.Completed;
FSteps[8].Children[1].Ready := FALSE;
FSteps[8].Children[1].Complete := TRUE;
FSteps[8].Children[1].Result := E_Result.Passed;
FSteps[8].Children[2].State := E_State.Completed;
FSteps[8].Children[2].Ready := FALSE;
FSteps[8].Children[2].Complete := TRUE;
FSteps[8].Children[2].Result := E_Result.Passed;
FSteps[8].Children[3].State := E_State.Completed;
FSteps[8].Children[3].Ready := FALSE;
FSteps[8].Children[3].Complete := TRUE;
FSteps[8].Children[3].Result := E_Result.Passed;
FSteps[8].ExpectedFinished := TRUE;
FSteps[8].ExpectedReleasedEntries[1] := 1;
FSteps[8].MaxActiveChildCount := 0;
{endregion}

{region "09 - Keep completion stable without further Starts"}
FSteps[9].Children[1].State := E_State.Completed;
FSteps[9].Children[1].Ready := FALSE;
FSteps[9].Children[1].Complete := TRUE;
FSteps[9].Children[1].Result := E_Result.Passed;
FSteps[9].Children[2].State := E_State.Completed;
FSteps[9].Children[2].Ready := FALSE;
FSteps[9].Children[2].Complete := TRUE;
FSteps[9].Children[2].Result := E_Result.Passed;
FSteps[9].Children[3].State := E_State.Completed;
FSteps[9].Children[3].Ready := FALSE;
FSteps[9].Children[3].Complete := TRUE;
FSteps[9].Children[3].Result := E_Result.Passed;
FSteps[9].ExpectedFinished := TRUE;
FSteps[9].MaxActiveChildCount := 0;
{endregion}
END_METHOD

END_FUNCTION_BLOCK

// ---- SelfTests/TestCases/TestSuite_ParallelOrchestration/Test_ParallelFirstFittingAdmission.TcPOU
{region 'Documentation'}
(*!
<summary>Skips a temporarily capacity-blocked same-slot child, starts fitting siblings, then admits the waiting child once.</summary>
<description>
Child 1 returns WaitingForCapacity twice while children 2 and 3 fit. All three later
overlap. Reservation responses test candidate selection only; real Event Buffer budget
arithmetic belongs to dedicated reservation tests.
</description>
*)
{endregion}
FUNCTION_BLOCK Test_ParallelFirstFittingAdmission EXTENDS OrchestrationTestBase

SUPER^();

{region 'Documentation'}
(*!
<summary>Defines independent per-cycle child responses and Parallel dispatch expectations.</summary>
*)
{endregion}
METHOD PROTECTED ConfigureScenario
FChildSlots[1] := 1;
FChildSlots[2] := 1;
FChildSlots[3] := 1;
FStepCount := 9;

{region "01 - Observe initial readiness"}
FSteps[1].Task := E_OrchestratorTask.Idle;
FSteps[1].ExpectedReady := TRUE;
{endregion}

{region "02 - Child 1 waits but child 2 fits"}
FSteps[2].Children[2].State := E_State.Running;
FSteps[2].Children[2].Ready := FALSE;
FSteps[2].ExecutionReservationResults[1] := E_EventReservationResult.WaitingForCapacity;
FSteps[2].ExpectedUnacceptedExecutionReservations[1] := 1;
FSteps[2].ExpectedStartChild := 2;
FSteps[2].ExpectedSlot := 1;
FSteps[2].ExpectedReservations[2] := 1;
FSteps[2].MaxActiveChildCount := 1;
{endregion}

{region "03 - Child 1 still waits but child 3 fits"}
FSteps[3].Children[2].State := E_State.Running;
FSteps[3].Children[2].Ready := FALSE;
FSteps[3].Children[3].State := E_State.Running;
FSteps[3].Children[3].Ready := FALSE;
FSteps[3].ExecutionReservationResults[1] := E_EventReservationResult.WaitingForCapacity;
FSteps[3].ExpectedUnacceptedExecutionReservations[1] := 1;
FSteps[3].ExpectedStartChild := 3;
FSteps[3].ExpectedSlot := 1;
FSteps[3].ExpectedReservations[2] := 1;
FSteps[3].ExpectedReservations[3] := 1;
FSteps[3].MaxActiveChildCount := 2;
{endregion}

{region "04 - Admit child 1 while its siblings remain active"}
FSteps[4].Children[1].State := E_State.Running;
FSteps[4].Children[1].Ready := FALSE;
FSteps[4].Children[2].State := E_State.Running;
FSteps[4].Children[2].Ready := FALSE;
FSteps[4].Children[3].State := E_State.Running;
FSteps[4].Children[3].Ready := FALSE;
FSteps[4].ExpectedStartChild := 1;
FSteps[4].ExpectedSlot := 1;
FSteps[4].ExpectedReservations[1] := 1;
FSteps[4].ExpectedReservations[2] := 1;
FSteps[4].ExpectedReservations[3] := 1;
FSteps[4].MaxActiveChildCount := 3;
{endregion}

{region "05 - Child 2 completes without interrupting its siblings"}
FSteps[5].Children[1].State := E_State.Running;
FSteps[5].Children[1].Ready := FALSE;
FSteps[5].Children[2].State := E_State.Completed;
FSteps[5].Children[2].Ready := FALSE;
FSteps[5].Children[2].Complete := TRUE;
FSteps[5].Children[2].Result := E_Result.Passed;
FSteps[5].Children[3].State := E_State.Running;
FSteps[5].Children[3].Ready := FALSE;
FSteps[5].ExpectedSlot := 1;
FSteps[5].ExpectedReservations[1] := 1;
FSteps[5].ExpectedReservations[2] := 1;
FSteps[5].ExpectedReservations[3] := 1;
FSteps[5].MaxActiveChildCount := 3;
{endregion}

{region "06 - Release child 2 then observe child 1 completion"}
FSteps[6].Children[1].State := E_State.Completed;
FSteps[6].Children[1].Ready := FALSE;
FSteps[6].Children[1].Complete := TRUE;
FSteps[6].Children[1].Result := E_Result.Passed;
FSteps[6].Children[2].State := E_State.Completed;
FSteps[6].Children[2].Ready := FALSE;
FSteps[6].Children[2].Complete := TRUE;
FSteps[6].Children[2].Result := E_Result.Passed;
FSteps[6].Children[3].State := E_State.Running;
FSteps[6].Children[3].Ready := FALSE;
FSteps[6].ExpectedSlot := 1;
FSteps[6].ExpectedReservations[1] := 1;
FSteps[6].ExpectedReservations[3] := 1;
FSteps[6].ExpectedReleasedEntries[2] := 1;
FSteps[6].MaxActiveChildCount := 2;
{endregion}

{region "07 - Release child 1 while child 3 completes"}
FSteps[7].Children[1].State := E_State.Completed;
FSteps[7].Children[1].Ready := FALSE;
FSteps[7].Children[1].Complete := TRUE;
FSteps[7].Children[1].Result := E_Result.Passed;
FSteps[7].Children[2].State := E_State.Completed;
FSteps[7].Children[2].Ready := FALSE;
FSteps[7].Children[2].Complete := TRUE;
FSteps[7].Children[2].Result := E_Result.Passed;
FSteps[7].Children[3].State := E_State.Completed;
FSteps[7].Children[3].Ready := FALSE;
FSteps[7].Children[3].Complete := TRUE;
FSteps[7].Children[3].Result := E_Result.Passed;
FSteps[7].ExpectedSlot := 1;
FSteps[7].ExpectedReservations[3] := 1;
FSteps[7].ExpectedReleasedEntries[1] := 1;
FSteps[7].MaxActiveChildCount := 1;
{endregion}

{region "08 - Finish only after child 3 reservation is released"}
FSteps[8].Children[1].State := E_State.Completed;
FSteps[8].Children[1].Ready := FALSE;
FSteps[8].Children[1].Complete := TRUE;
FSteps[8].Children[1].Result := E_Result.Passed;
FSteps[8].Children[2].State := E_State.Completed;
FSteps[8].Children[2].Ready := FALSE;
FSteps[8].Children[2].Complete := TRUE;
FSteps[8].Children[2].Result := E_Result.Passed;
FSteps[8].Children[3].State := E_State.Completed;
FSteps[8].Children[3].Ready := FALSE;
FSteps[8].Children[3].Complete := TRUE;
FSteps[8].Children[3].Result := E_Result.Passed;
FSteps[8].ExpectedFinished := TRUE;
FSteps[8].ExpectedReleasedEntries[3] := 1;
FSteps[8].MaxActiveChildCount := 0;
{endregion}

{region "09 - No skipped child or repeated Start remains"}
FSteps[9].Children[1].State := E_State.Completed;
FSteps[9].Children[1].Ready := FALSE;
FSteps[9].Children[1].Complete := TRUE;
FSteps[9].Children[1].Result := E_Result.Passed;
FSteps[9].Children[2].State := E_State.Completed;
FSteps[9].Children[2].Ready := FALSE;
FSteps[9].Children[2].Complete := TRUE;
FSteps[9].Children[2].Result := E_Result.Passed;
FSteps[9].Children[3].State := E_State.Completed;
FSteps[9].Children[3].Ready := FALSE;
FSteps[9].Children[3].Complete := TRUE;
FSteps[9].Children[3].Result := E_Result.Passed;
FSteps[9].ExpectedFinished := TRUE;
FSteps[9].MaxActiveChildCount := 0;
{endregion}
END_METHOD

END_FUNCTION_BLOCK

// ---- SelfTests/TestCases/TestSuite_ParallelOrchestration/Test_ParallelMissingStartReaction.TcPOU
{region 'Documentation'}
(*!
<summary>Rejects a missing same-slot Start reaction without releasing a running sibling's reservation or starting another child.</summary>
<description>
Child 1 runs when child 2 ignores Start and stays Idle. The following helper call must
release only child 2 and hold one isolated Framework diagnostic. Child 1 subsequently
completes naturally; child 3 must never receive Start.
</description>
*)
{endregion}
FUNCTION_BLOCK Test_ParallelMissingStartReaction EXTENDS OrchestrationTestBase

SUPER^();

{region 'Documentation'}
(*!
<summary>Defines independent per-cycle child responses and Parallel dispatch expectations.</summary>
*)
{endregion}
METHOD PROTECTED ConfigureScenario
FChildSlots[1] := 1;
FChildSlots[2] := 1;
FChildSlots[3] := 1;
FStepCount := 8;

{region "01 - Observe initial readiness"}
FSteps[1].Task := E_OrchestratorTask.Idle;
FSteps[1].ExpectedReady := TRUE;
{endregion}

{region "02 - Start child 1 normally"}
FSteps[2].Children[1].State := E_State.Running;
FSteps[2].Children[1].Ready := FALSE;
FSteps[2].ExpectedStartChild := 1;
FSteps[2].ExpectedSlot := 1;
FSteps[2].ExpectedReservations[1] := 1;
FSteps[2].MaxActiveChildCount := 1;
{endregion}

{region "03 - Request child 2 Start but keep it Idle"}
FSteps[3].Children[1].State := E_State.Running;
FSteps[3].Children[1].Ready := FALSE;
FSteps[3].ExpectedStartChild := 2;
FSteps[3].ExpectedSlot := 1;
FSteps[3].ExpectedReservations[1] := 1;
FSteps[3].ExpectedReservations[2] := 1;
FSteps[3].MaxActiveChildCount := 2;
{endregion}

{region "04 - Reject child 2 while retaining child 1 reservation"}
FSteps[4].Children[1].State := E_State.Running;
FSteps[4].Children[1].Ready := FALSE;
FSteps[4].ExpectedSlot := 1;
FSteps[4].ExpectedReservations[1] := 1;
FSteps[4].ExpectedReleasedEntries[2] := 1;
FSteps[4].MaxActiveChildCount := 1;
FSteps[4].ExpectedResult := E_Result.Error;
FSteps[4].ExpectedDiagnosticCount := 1;
{endregion}

{region "05 - Hold the error without retry or child 3 Start"}
FSteps[5].Children[1].State := E_State.Running;
FSteps[5].Children[1].Ready := FALSE;
FSteps[5].ExpectedSlot := 1;
FSteps[5].ExpectedReservations[1] := 1;
FSteps[5].MaxActiveChildCount := 1;
FSteps[5].ExpectedResult := E_Result.Error;
FSteps[5].ExpectedDiagnosticCount := 1;
{endregion}

{region "06 - Child 1 finishes independently of the held helper error"}
FSteps[6].Children[1].State := E_State.Completed;
FSteps[6].Children[1].Ready := FALSE;
FSteps[6].Children[1].Complete := TRUE;
FSteps[6].Children[1].Result := E_Result.Passed;
FSteps[6].ExpectedSlot := 1;
FSteps[6].ExpectedReservations[1] := 1;
FSteps[6].MaxActiveChildCount := 1;
FSteps[6].ExpectedResult := E_Result.Error;
FSteps[6].ExpectedDiagnosticCount := 1;
{endregion}

{region "07 - Release child 1 only after terminal observation"}
FSteps[7].Children[1].State := E_State.Completed;
FSteps[7].Children[1].Ready := FALSE;
FSteps[7].Children[1].Complete := TRUE;
FSteps[7].Children[1].Result := E_Result.Passed;
FSteps[7].ExpectedSlot := 1;
FSteps[7].ExpectedReleasedEntries[1] := 1;
FSteps[7].MaxActiveChildCount := 0;
FSteps[7].ExpectedResult := E_Result.Error;
FSteps[7].ExpectedDiagnosticCount := 1;
{endregion}

{region "08 - Keep the error without repeated diagnostics or Starts"}
FSteps[8].Children[1].State := E_State.Completed;
FSteps[8].Children[1].Ready := FALSE;
FSteps[8].Children[1].Complete := TRUE;
FSteps[8].Children[1].Result := E_Result.Passed;
FSteps[8].ExpectedSlot := 1;
FSteps[8].MaxActiveChildCount := 0;
FSteps[8].ExpectedResult := E_Result.Error;
FSteps[8].ExpectedDiagnosticCount := 1;
{endregion}
END_METHOD

END_FUNCTION_BLOCK

// ---- SelfTests/TestCases/TestSuite_ParallelOrchestration/Test_ParallelReadinessLost.TcPOU
{region 'Documentation'}
(*!
<summary>Detects a same-slot child's readiness loss after valid admission and prevents further Starts.</summary>
<description>
All children initially report ready. Child 2 loses readiness while child 1 starts, as when
a shared resource changes. Child 1 may finish, but neither unstarted child is dispatched
and one diagnostic remains held.
</description>
*)
{endregion}
FUNCTION_BLOCK Test_ParallelReadinessLost EXTENDS OrchestrationTestBase

SUPER^();

{region 'Documentation'}
(*!
<summary>Defines reachable child responses and independent per-cycle expectations.</summary>
*)
{endregion}
METHOD PROTECTED ConfigureScenario
FChildSlots[1] := 1;
FChildSlots[2] := 1;
FChildSlots[3] := 1;
FStepCount := 8;

{region "01 - Observe initial group readiness"}
FSteps[1].Task := E_OrchestratorTask.Idle;
FSteps[1].ExpectedReady := TRUE;
{endregion}

{region "02 - Start child 1 while child 2 loses readiness"}
FSteps[2].Children[1].State := E_State.Running;
FSteps[2].Children[1].Ready := FALSE;
FSteps[2].Children[2].State := E_State.Idle;
FSteps[2].Children[2].Ready := FALSE;
FSteps[2].ExpectedStartChild := 1;
FSteps[2].ExpectedSlot := 1;
FSteps[2].ExpectedReservations[1] := 1;
FSteps[2].MaxActiveChildCount := 1;
{endregion}

{region "03 - Detect lost readiness before another Start"}
FSteps[3].Children[1].State := E_State.Running;
FSteps[3].Children[1].Ready := FALSE;
FSteps[3].Children[2].State := E_State.Idle;
FSteps[3].Children[2].Ready := FALSE;
FSteps[3].ExpectedSlot := 1;
FSteps[3].ExpectedReservations[1] := 1;
FSteps[3].MaxActiveChildCount := 1;
FSteps[3].ExpectedResult := E_Result.Error;
FSteps[3].ExpectedDiagnosticCount := 1;
{endregion}

{region "04 - Keep the active child reserved without redispatch"}
FSteps[4].Children[1].State := E_State.Running;
FSteps[4].Children[1].Ready := FALSE;
FSteps[4].Children[2].State := E_State.Idle;
FSteps[4].Children[2].Ready := FALSE;
FSteps[4].ExpectedSlot := 1;
FSteps[4].ExpectedReservations[1] := 1;
FSteps[4].MaxActiveChildCount := 1;
FSteps[4].ExpectedResult := E_Result.Error;
FSteps[4].ExpectedDiagnosticCount := 1;
{endregion}

